      movej([-1.2302089344500047, -1.2969853503591224, -1.875639182904262, -1.539621866126728, 1.5731943360401213, -2.80099559440227], a=1.3962634015954636, v=1.0471975511965976)
    elif (32 == switch_1):
      $ 1983 "Case 32"
      $ 1985 "decap_Vial"
      $ 1986 "Set GRP_3F_Open=On"
      set_standard_digital_out(5, True)
      $ 1987 "MoveJ"
      $ 1988 "Waypoint_87" "breakAfter"
      movej(get_inverse_kin(Waypoint_87_p, qnear=Waypoint_87_q), a=0.5235987755982988, v=0.4363323129985824)
      $ 1989 "MoveL"
      $ 1990 "Vial_3FG_plac_1" "breakAfter"
      movel(Vial_3FG_plac_1_p, a=0.5, v=0.1)
      $ 1991 "Set GRP_3F_Open=Off"
      set_standard_digital_out(5, False)
      $ 1992 "Wait: 0.5"
      sleep(0.5)
      $ 1993 "MoveL"
      $ 1994 "Waypoint_88" "breakAfter"
      movel(Waypoint_88_p, a=0.5, v=0.1, r=0.05)
      $ 1995 "MoveJ"
      $ 1996 "cap_dump_1" "breakAfter"
      movej(get_inverse_kin(cap_dump_1_p, qnear=cap_dump_1_q), a=0.5235987755982988, v=0.4363323129985824)
      # begin: URCap Program Node
      #   Source: Robotiq_Grippers, 3.17.0.105337, Robotiq Inc.
      #   Type: Gripper
      $ 1997 "Gripper Open (1)"
      if not(gripper_connected[0]):
        popup("Gripper 1 must be connected to run this program.", "No connection", False, True, True)
      end
      if not(rq_is_gripper_activated("1")):
        popup("Gripper 1 is not activated. Go to Installation tab > Gripper to activate it and run the program again.", "Not activated", False, True, True)
      end
      rq_set_pos_spd_for(0, 255, 255, "1")
      rq_wait_pos_spe_for_request(0, 255, 255, "1")
      rq_go_to("1")
      rq_wait("1")
      # end: URCap Program Node
      $ 1998 "MoveJ"
      $ 1999 "Waypoint_89" "breakAfter"
      movej(get_inverse_kin(Waypoint_89_p, qnear=Waypoint_89_q), a=0.5235987755982988, v=0.4363323129985824, r=0.05)
      $ 2000 "MoveL"
      $ 2001 "Vial_3FG_plac_2" "breakAfter"
      movel(Vial_3FG_plac_2_p, a=0.5, v=0.1)
      # begin: URCap Program Node
      #   Source: Robotiq_Grippers, 3.17.0.105337, Robotiq Inc.
      #   Type: Gripper
      $ 2002 "Gripper Close (1)"
      if not(gripper_connected[0]):
        popup("Gripper 1 must be connected to run this program.", "No connection", False, True, True)
      end
      if not(rq_is_gripper_activated("1")):
        popup("Gripper 1 is not activated. Go to Installation tab > Gripper to activate it and run the program again.", "Not activated", False, True, True)
      end
      rq_set_pos_spd_for(255, 204, 255, "1")
      rq_wait_pos_spe_for_request(255, 204, 255, "1")
      rq_go_to("1")
      rq_wait("1")
      # end: URCap Program Node
      $ 2009 "Decap"
      $ 2010 "Action_Info≔'decapping'"
      global Action_Info="decapping"
      $ 2011 "Set GRP_3F_Enable=On"
      set_standard_digital_out(4, True)
      $ 2012 "Set GRP_3F_Decap=On"
      set_standard_digital_out(3, True)
      $ 2013 "Force"
      sleep(0.02)
      zero_ftsensor()
      force_mode(p[0.0,0.0,0.0,0.0,0.0,0.0], [0, 0, 1, 0, 0, 0], [0.0, 0.0, 1.0, 0.0, 0.0, 0.0], 2, [0.1, 0.1, 0.001, 0.3490658503988659, 0.3490658503988659, 0.3490658503988659])
      $ 2014 "check_decapping(offset=0.015, timeout=10, abort=CMD_Hold)" "noBreak"
      check_decapping(offset=0.015, timeout=10, abort=CMD_Hold)
      end_force_mode()
      stopl(5.0)
      $ 2015 "Set GRP_3F_Decap=Off"
      set_standard_digital_out(3, False)
      $ 2016 "Set GRP_3F_Enable=Off"
      set_standard_digital_out(4, False)
      $ 2017 "MoveL"
      $ 2018 "Waypoint_90" "breakAfter"
      movel(Waypoint_90_p, a=0.5, v=0.1, r=0.05)
      $ 2019 "MoveJ"
      $ 2020 "cap_dump_2" "breakAfter"
      movej(get_inverse_kin(cap_dump_2_p, qnear=cap_dump_2_q), a=0.5235987755982988, v=0.4363323129985824)
      # begin: URCap Program Node
      #   Source: Robotiq_Grippers, 3.17.0.105337, Robotiq Inc.
      #   Type: Gripper
      $ 2021 "Gripper Open (1)"
      if not(gripper_connected[0]):
        popup("Gripper 1 must be connected to run this program.", "No connection", False, True, True)
      end
      if not(rq_is_gripper_activated("1")):
        popup("Gripper 1 is not activated. Go to Installation tab > Gripper to activate it and run the program again.", "Not activated", False, True, True)
      end
      rq_set_pos_spd_for(0, 204, 255, "1")
      rq_wait_pos_spe_for_request(0, 204, 255, "1")
      rq_go_to("1")
      rq_wait("1")
      # end: URCap Program Node
      $ 2022 "MoveJ"
      $ 2023 "Waypoint_91" "breakAfter"
      movej(get_inverse_kin(Waypoint_91_p, qnear=Waypoint_91_q), a=0.5235987755982988, v=0.4363323129985824, r=0.036)
    elif (33 == switch_1):
      $ 2024 "Case 33"
      $ 2025 "Shake and liquid transfer"
      $ 2026 "MoveL"
      $ 2027 "Vial_liq_abov_1" "breakAfter"
      movel(Vial_liq_abov_1_p, a=0.5, v=0.1)
      $ 2028 "Vial_liq_pick_3" "breakAfter"
      movel(Vial_liq_pick_3_p, a=0.5, v=0.1)
      $ 2029 "Vial_liq_pick_4" "breakAfter"
      movel(Vial_liq_pick_4_p, a=0.5, v=0.1)
      # begin: URCap Program Node
      #   Source: Robotiq_Grippers, 3.17.0.105337, Robotiq Inc.
      #   Type: Gripper
      $ 2030 "Gripper Close (1)"
      if not(gripper_connected[0]):
        popup("Gripper 1 must be connected to run this program.", "No connection", False, True, True)
      end
      if not(rq_is_gripper_activated("1")):
        popup("Gripper 1 is not activated. Go to Installation tab > Gripper to activate it and run the program again.", "Not activated", False, True, True)
      end
      rq_set_pos_spd_for(255, 82, 71, "1")
      rq_wait_pos_spe_for_request(255, 82, 71, "1")
      rq_go_to("1")
      rq_wait("1")
      # end: URCap Program Node
      $ 2031 "Wait: 1.0"
      sleep(1.0)
      $ 2032 "Set GRP_3F_Open=On"
      set_standard_digital_out(5, True)
      $ 2033 "Wait: 0.5"
      sleep(0.5)
      $ 2034 "Vial_liq_abov_2" "breakAfter"
      movel(Vial_liq_abov_2_p, a=0.3, v=0.05, r=0.05)
      $ 2035 "MoveL"
      $ 2036 "Liquid_midway_1" "breakAfter"
      movel(Liquid_midway_1_p, a=0.5, v=0.1)
      $ 2037 "Loop 3 times"
      Loop_1 = 0
      while (Loop_1 < 3):
        $ 2038 "shake_3" "breakAfter"
        movel(shake_3_p, a=2.0, v=0.5)
        $ 2039 "shake_4" "breakAfter"
        movel(shake_4_p, a=2.0, v=0.5)
        Loop_1 = Loop_1 + 1
      end
      $ 2040 "drop_above_3" "breakAfter"
      movel(drop_above_3_p, a=0.5, v=0.1)
      $ 2041 "drop_above_4" "breakAfter"
      movel(drop_above_4_p, a=0.5, v=0.1)
      $ 2042 "liq_tran_3" "breakAfter"
      movel(liq_tran_3_p, a=0.5, v=0.05, r=0.008)
      $ 2043 "Wait: 1.0"
      sleep(1.0)
      $ 2044 "drop_above_5" "breakAfter"
      movel(drop_above_5_p, a=0.5, v=0.1)
      $ 2045 "Waypoint_92" "breakAfter"
      movel(Waypoint_92_p, a=0.5, v=0.1)
      $ 2046 "liq_tran_4" "breakAfter"
      movel(liq_tran_4_p, a=0.5, v=0.05)
      $ 2047 "Wait: 1.0"
      sleep(1.0)
      $ 2048 "drop_above_6" "breakAfter"
      movel(drop_above_6_p, a=0.5, v=0.1)
      $ 2049 "drop_above_7" "breakAfter"
      movel(drop_above_7_p, a=0.5, v=0.1)
      $ 2050 "Liquid_midway_2" "breakAfter"
      movel(Liquid_midway_2_p, a=0.5, v=0.1)
      $ 2051 "MoveL"
      $ 2052 "Vial_drop_abo_1" "breakAfter"
      movel(Vial_drop_abo_1_p, a=0.5, v=0.1)
      $ 2053 "Vial_liq_drop_1" "breakAfter"
      movel(Vial_liq_drop_1_p, a=0.5, v=0.1)
      # begin: URCap Program Node
      #   Source: Robotiq_Grippers, 3.17.0.105337, Robotiq Inc.
      #   Type: Gripper
      $ 2054 "Gripper Open (1)"
      if not(gripper_connected[0]):
        popup("Gripper 1 must be connected to run this program.", "No connection", False, True, True)
      end
      if not(rq_is_gripper_activated("1")):
        popup("Gripper 1 is not activated. Go to Installation tab > Gripper to activate it and run the program again.", "Not activated", False, True, True)
      end
      rq_set_pos_spd_for(0, 82, 71, "1")
      rq_wait_pos_spe_for_request(0, 82, 71, "1")
      rq_go_to("1")
      rq_wait("1")
      # end: URCap Program Node
      $ 2055 "Vial_drop_abo_2" "breakAfter"
      movel(Vial_drop_abo_2_p, a=0.5, v=0.1)
    elif (34 == switch_1):
      $ 2056 "Case 34"
      $ 2057 "Task≔'Dosing'"
      global Task="Dosing"
      $ 2058 "Powder dosing all"
      $ 2059 "send_target_info()"
      send_target_info()
      $ 2060 "zero_scale()"
      zero_scale()
      $ 2061 "prev_spat≔''"
      global prev_spat=""
      $ 2062 "spatula≔''"
      global spatula=""
      $ 2063 "send_powder_info()"
      send_powder_info()
      $ 2064 "Set AO[0]=0.0"
      set_standard_analog_out(0, 0.0)
      $ 2065 "Wait: 0.2"
      sleep(0.2)
      $ 2066 "reach pots decapping pose"
      # begin: URCap Program Node
      #   Source: SensoPart VISOR Robotic, 2.0.6, SensoPart Industriesensorik GmbH
      #   Type: VISOR Robotic App
      $ 2072 "VISOR Easy Pick"
      def visorFuncEasyPick_a93150():
        # begin: URCap Program Node
        #   Source: SensoPart VISOR Robotic, 2.0.6, SensoPart Industriesensorik GmbH
        #   Type: Easy Pick Setup
        $ 2073 "# 1 Setup" "noBreak"
        local easyPickVisorId = 1
        local easyPickArmMounted = True
        local easyPickSetJob = True
        local easyPickJobName = "Weight_scale"
        local easyPickAtImgAcq = False
        local easyPickImgAcqPose = Trigger
        # end: URCap Program Node
        # begin: URCap Program Node
        #   Source: SensoPart VISOR Robotic, 2.0.6, SensoPart Industriesensorik GmbH
        #   Type: Process
        $ 2074 "Process" "noBreak"
        local easyPickObjTaken = False
        local easyPickTrigger = False
        local easyPickPoseIdx = 0
        local easyPickPose = p[0,0,0,0,0,0]
        def easyPickFuncTrigger(visorId, setJob, jobName, arm):
        if (setJob):
          visor_changeJob(visorId, jobName, 6000)
        end
        if (arm):
          visor_trigger(visorId, 6000, "arm")
        else:
          visor_trigger(visorId, 6000)
        end
        global easyPickParts_4=visor_partsFound(visorId)
        visor_easyPickUpdate(visorId, "parts", visor_partsFound(visorId))
        return visor_getPose3d(visorId, 0)
      end
      while (not easyPickObjTaken):
        easyPickTrigger = (easyPickCount_4 >= visor_partsFound(easyPickVisorId)) or (easyPickCount_4 > 9) or (not visor_easyPickCheckIdent("3d2ec7", easyPickVisorId))
        if (easyPickTrigger):
          easyPickCount_4 = 0
        end
        easyPickPoseIdx = easyPickCount_4
        easyPickPose = visor_getPose3d(easyPickVisorId, easyPickPoseIdx)
        visor_easyPickUpdate(easyPickVisorId, "counter", easyPickPoseIdx)
        # begin: URCap Program Node
        #   Source: SensoPart VISOR Robotic, 2.0.6, SensoPart Industriesensorik GmbH
        #   Type: Image Acquisition Pose
        $ 2075 "Image Acquisition Pose" "noBreak"
        if (easyPickTrigger):
          if (not easyPickAtImgAcq):
            movej(pose_trans(easyPickImgAcqPose,p[0.0000,0.0000,-0.0000,0.0000,0.0000,0.0000]),a=1.3963,v=1.0472,t=0.000000,r=0.000000)
            easyPickAtImgAcq = True
          end
          easyPickPose = easyPickFuncTrigger(easyPickVisorId, easyPickSetJob, easyPickJobName, easyPickArmMounted)
        end
        # end: URCap Program Node
        # begin: URCap Program Node
        #   Source: SensoPart VISOR Robotic, 2.0.6, SensoPart Industriesensorik GmbH
        #   Type: Object Detected
        $ 2076 "Object Detected" "noBreak"
        if (visor_partsFound(easyPickVisorId) > 0):
          $ 2077 "Open Gripper" "noBreak"
          $ 2078 "weight_value≔get_weight()" "noBreak"
          global weight_value=get_weight()
          $ 2079 "Wait: 1.0" "noBreak"
          sleep(1.0)
          $ 2080 "diff≔target_weight-weight_value" "noBreak"
          global diff=target_weight-weight_value
          $ 2081 "compute_level_percent(W_now, weight_value)" "noBreak"
          compute_level_percent(W_now, weight_value)
          $ 2082 "send_level_info()" "noBreak"
          send_level_info()
          $ 2083 "spatula≔select_spatula(Flowability, level, diff, bulk_density, mouth_d)" "noBreak"
          global spatula=select_spatula(Flowability, level, diff, bulk_density, mouth_d)
          $ 2084 "Wait: 0.2" "noBreak"
          sleep(0.2)
          $ 2085 "send_spatula_info()" "noBreak"
          send_spatula_info()
          $ 2086 "If spatula ≟ 'spatula_L'" "noBreak"
          if (spatula  ==  "spatula_L"):
            $ 2087 "MoveJ" "noBreak"
            $ 2088 "Spatula_otw" "noBreak"
            movej(get_inverse_kin(Spatula_otw_p, qnear=Spatula_otw_q), a=1.3962634015954636, v=1.0471975511965976)
            $ 2089 "pick_spat_L_abv" "noBreak"
            movej(get_inverse_kin(pick_spat_L_abv_p, qnear=pick_spat_L_abv_q), a=1.3962634015954636, v=1.0471975511965976)
            $ 2090 "MoveL" "noBreak"
            $ 2091 "spat_L_pick" "noBreak"
            movel(spat_L_pick_p, a=1.2, v=0.25)
            # begin: URCap Program Node
            #   Source: Robotiq_Grippers, 3.17.0.105337, Robotiq Inc.
            #   Type: Gripper
            $ 2092 "Gripper Close (1)" "noBreak"
            if not(gripper_connected[0]):
              popup("Gripper 1 must be connected to run this program.", "No connection", False, True, True)
            end
            if not(rq_is_gripper_activated("1")):
              popup("Gripper 1 is not activated. Go to Installation tab > Gripper to activate it and run the program again.", "Not activated", False, True, True)
            end
            rq_set_pos_spd_for(255, 0, 77, "1")
            rq_wait_pos_spe_for_request(255, 0, 77, "1")
            rq_go_to("1")
            rq_wait("1")
            # end: URCap Program Node
            $ 2093 "spat_L_lift" "noBreak"
            movel(spat_L_lift_p, a=1.2, v=0.25, r=0.01)
            $ 2094 "spat_L_side" "noBreak"
            movel(spat_L_side_p, a=1.2, v=0.25, r=0.01)
            $ 2095 "spat_L_up" "noBreak"
            movel(spat_L_up_p, a=1.2, v=0.25, r=0.05)
            $ 2096 "MoveJ" "noBreak"
            $ 2097 "Spatula_otw" "noBreak"
            movej(get_inverse_kin(Spatula_otw_p, qnear=Spatula_otw_q), a=1.3962634015954636, v=1.0471975511965976)
          else:
            $ 2098 "ElseIf spatula ≟'spatula_M'" "noBreak"
            if (spatula  == "spatula_M"):
              $ 2099 "MoveJ" "noBreak"
              $ 2100 "Spatula_otw" "noBreak"
              movej(get_inverse_kin(Spatula_otw_p, qnear=Spatula_otw_q), a=1.3962634015954636, v=1.0471975511965976)
              $ 2101 "spat_M_up" "noBreak"
              movej(get_inverse_kin(spat_M_up_p, qnear=spat_M_up_q), a=1.3962634015954636, v=1.0471975511965976, r=0.05)
              $ 2102 "MoveL" "noBreak"
              $ 2103 "spat_M_pick" "noBreak"
              movel(spat_M_pick_p, a=1.2, v=0.25)
              # begin: URCap Program Node
              #   Source: Robotiq_Grippers, 3.17.0.105337, Robotiq Inc.
              #   Type: Gripper
              $ 2104 "Gripper Close (1)" "noBreak"
              if not(gripper_connected[0]):
                popup("Gripper 1 must be connected to run this program.", "No connection", False, True, True)
              end
              if not(rq_is_gripper_activated("1")):
                popup("Gripper 1 is not activated. Go to Installation tab > Gripper to activate it and run the program again.", "Not activated", False, True, True)
              end
              rq_set_pos_spd_for(255, 0, 77, "1")
              rq_wait_pos_spe_for_request(255, 0, 77, "1")
              rq_go_to("1")
              rq_wait("1")
              # end: URCap Program Node
              $ 2105 "spat_M_up" "noBreak"
              movel(spat_M_up_p, a=1.2, v=0.25, r=0.05)
              $ 2106 "Spatula_otw" "noBreak"
              movel(Spatula_otw_p, a=1.2, v=0.25)
              $ 2107 "switch_spat_M≔ False " "noBreak"
              global switch_spat_M=  False
            else:
              $ 2108 "ElseIf spatula≟'spatula_S'" "noBreak"
              if (spatula == "spatula_S"):
                $ 2109 "MoveJ" "noBreak"
                $ 2110 "Spatula_otw" "noBreak"
                movej(get_inverse_kin(Spatula_otw_p, qnear=Spatula_otw_q), a=1.3962634015954636, v=1.0471975511965976)
                $ 2111 "spat_S_Up_7" "noBreak"
                movej(get_inverse_kin(spat_S_Up_7_p, qnear=spat_S_Up_7_q), a=1.3962634015954636, v=1.0471975511965976, r=0.05)
                $ 2112 "MoveL" "noBreak"
                $ 2113 "spat_S_Pick_4" "noBreak"
                movel(spat_S_Pick_4_p, a=1.2, v=0.25)
                # begin: URCap Program Node
                #   Source: Robotiq_Grippers, 3.17.0.105337, Robotiq Inc.
                #   Type: Gripper
                $ 2114 "Gripper Close (1)" "noBreak"
                if not(gripper_connected[0]):
                  popup("Gripper 1 must be connected to run this program.", "No connection", False, True, True)
                end
                if not(rq_is_gripper_activated("1")):
                  popup("Gripper 1 is not activated. Go to Installation tab > Gripper to activate it and run the program again.", "Not activated", False, True, True)
                end
                rq_set_pos_spd_for(255, 0, 77, "1")
                rq_wait_pos_spe_for_request(255, 0, 77, "1")
                rq_go_to("1")
                rq_wait("1")
                # end: URCap Program Node
                $ 2115 "spat_S_Up_8" "noBreak"
                movel(spat_S_Up_8_p, a=1.2, v=0.25, r=0.05)
                $ 2116 "Spatula_otw" "noBreak"
                movel(Spatula_otw_p, a=1.2, v=0.25)
                $ 2117 "switch_spat_S≔ False " "noBreak"
                global switch_spat_S=  False
              else:
                $ 2118 "ElseIf spatula≟'spatula_flat_M'" "noBreak"
                if (spatula == "spatula_flat_M"):
                  $ 2119 "MoveJ" "noBreak"
                  $ 2120 "Spatula_otw" "noBreak"
                  movej(get_inverse_kin(Spatula_otw_p, qnear=Spatula_otw_q), a=1.3962634015954636, v=1.0471975511965976)
                  $ 2121 "spat_flatM_up" "noBreak"
                  movej(get_inverse_kin(spat_flatM_up_p, qnear=spat_flatM_up_q), a=1.3962634015954636, v=1.0471975511965976, r=0.05)
                  $ 2122 "MoveL" "noBreak"
                  $ 2123 "spat_flatM_pick" "noBreak"
                  movel(spat_flatM_pick_p, a=1.2, v=0.25)
                  # begin: URCap Program Node
                  #   Source: Robotiq_Grippers, 3.17.0.105337, Robotiq Inc.
                  #   Type: Gripper
                  $ 2124 "Gripper Close (1)" "noBreak"
                  if not(gripper_connected[0]):
                    popup("Gripper 1 must be connected to run this program.", "No connection", False, True, True)
                  end
                  if not(rq_is_gripper_activated("1")):
                    popup("Gripper 1 is not activated. Go to Installation tab > Gripper to activate it and run the program again.", "Not activated", False, True, True)
                  end
                  rq_set_pos_spd_for(255, 0, 77, "1")
                  rq_wait_pos_spe_for_request(255, 0, 77, "1")
                  rq_go_to("1")
                  rq_wait("1")
                  # end: URCap Program Node
                  $ 2125 "spat_flatM_up" "noBreak"
                  movel(spat_flatM_up_p, a=1.2, v=0.25, r=0.05)
                  $ 2126 "Spatula_otw" "noBreak"
                  movel(Spatula_otw_p, a=1.2, v=0.25)
                  $ 2127 "switch_spat_F_M≔ False " "noBreak"
                  global switch_spat_F_M=  False
                else:
                  $ 2128 "ElseIf spatula≟'spatula_flat_S'" "noBreak"
                  if (spatula == "spatula_flat_S"):
                    $ 2129 "MoveJ" "noBreak"
                    $ 2130 "Spatula_otw" "noBreak"
                    movej(get_inverse_kin(Spatula_otw_p, qnear=Spatula_otw_q), a=1.3962634015954636, v=1.0471975511965976)
                    $ 2131 "spat_flatS_up" "noBreak"
                    movej(get_inverse_kin(spat_flatS_up_p, qnear=spat_flatS_up_q), a=1.3962634015954636, v=1.0471975511965976, r=0.05)
                    $ 2132 "MoveL" "noBreak"
                    $ 2133 "spat_flatS_pick" "noBreak"
                    movel(spat_flatS_pick_p, a=1.2, v=0.25)
                    # begin: URCap Program Node
                    #   Source: Robotiq_Grippers, 3.17.0.105337, Robotiq Inc.
                    #   Type: Gripper
                    $ 2134 "Gripper Close (1)" "noBreak"
                    if not(gripper_connected[0]):
                      popup("Gripper 1 must be connected to run this program.", "No connection", False, True, True)
                    end
                    if not(rq_is_gripper_activated("1")):
                      popup("Gripper 1 is not activated. Go to Installation tab > Gripper to activate it and run the program again.", "Not activated", False, True, True)
                    end
                    rq_set_pos_spd_for(255, 0, 77, "1")
                    rq_wait_pos_spe_for_request(255, 0, 77, "1")
                    rq_go_to("1")
                    rq_wait("1")
                    # end: URCap Program Node
                    $ 2135 "spat_flatS_up" "noBreak"
                    movel(spat_flatS_up_p, a=1.2, v=0.25, r=0.05)
                    $ 2136 "Spatula_otw" "noBreak"
                    movel(Spatula_otw_p, a=1.2, v=0.25)
                    $ 2137 "switch_spat_F_S≔ False " "noBreak"
                    global switch_spat_F_S=  False
                  end
                end
              end
            end
          end
          $ 2138 "Action_Info≔'Scooping'" "noBreak"
          global Action_Info="Scooping"
          $ 2139 "auto_tilt_and_scoop(W_now, target_weight, weight_value)" "noBreak"
          auto_tilt_and_scoop(W_now, target_weight, weight_value)
          $ 2140 "Action_Info≔'Dosing'" "noBreak"
          global Action_Info="Dosing"
          # begin: URCap Program Node
          #   Source: SensoPart VISOR Robotic, 2.0.6, SensoPart Industriesensorik GmbH
          #   Type: Approach Pose
          $ 2141 "Approach Pose" "noBreak"
          movej(pose_trans(easyPickPose,p[0.0000,0.0000,-0.0000,0.0000,0.0000,0.0000]),a=0.2618,v=0.1745,t=0.000000,r=0.000000)
          # end: URCap Program Node
          # begin: URCap Program Node
          #   Source: SensoPart VISOR Robotic, 2.0.6, SensoPart Industriesensorik GmbH
          #   Type: Target Pose
          $ 2142 "Target Pose" "noBreak"
          movel(pose_trans(easyPickPose,p[0.0000,0.0000,-0.0000,0.0000,0.0000,0.0000]),a=0.0500,v=0.0200,t=0.000000,r=0.000000)
          # end: URCap Program Node
          $ 2143 "Close Gripper" "noBreak"
          $ 2144 "dispense_pos≔get_actual_tcp_pose()" "noBreak"
          global dispense_pos= get_actual_tcp_pose ()
          $ 2145 "Loop weight_value≤target_weight " "noBreak"
          thread Thread_while_2145():
            while (True):
              $ 2146 "MoveL" "noBreak"
              $ 2147 "dispense_pos" "noBreak"
              movel(dispense_pos, a=0.2, v=0.1)
              $ 2148 "log_weight()" "noBreak"
              log_weight()
              $ 2149 "If level≥85" "noBreak"
              if (level >= 85):
                $ 2150 "Rotate()" "noBreak"
                Rotate()
              end
              $ 2151 "If level≤85" "noBreak"
              if (level <= 85):
                $ 2152 "tilt_to_home()" "noBreak"
                tilt_to_home()
              end
              $ 2153 "Start_thread≔ True " "noBreak"
              global Start_thread=  True
              $ 2154 "vib_thread≔ True " "noBreak"
              global vib_thread=  True
              $ 2155 "Wait: 0.5" "noBreak"
              sleep(0.5)
              $ 2156 "If diff ≥(target_g*1.1)" "noBreak"
              if (diff  >= (target_g*1.1)):
                $ 2157 "tilt_pose≔pose_trans(get_actual_tcp_pose(), p[0, 0, 0, 0, 0, 2.0])" "noBreak"
                global tilt_pose=pose_trans(get_actual_tcp_pose(), p[0, 0, 0, 0, 0, 2.0])
                $ 2158 "movel(tilt_pose, a=0.5, v=0.5, r=0.00001)" "noBreak"
                movel(tilt_pose, a=0.5, v=0.5, r=0.00001)
              else:
                $ 2159 "Else" "noBreak"
                $ 2160 "Loop weight_value≤(target_weight-0.00) and tilt_angle≥(-1.999) and tilt_angle≤0.5" "noBreak"
                thread Thread_while_2160():
                  while (True):
                    $ 2161 "current_error≔target_weight-weight_value" "noBreak"
                    global current_error=target_weight-weight_value
                    $ 2162 "Integral_error≔Integral_error+current_error*dt" "noBreak"
                    global Integral_error=Integral_error+current_error*dt
                    $ 2163 "derivative≔(current_error-previous_error)/dt" "noBreak"
                    global derivative=(current_error-previous_error)/dt
                    $ 2164 "tilt_increment≔(kp*current_error)+(ki*Integral_error)+(kd*derivative)" "noBreak"
                    global tilt_increment=(kp*current_error)+(ki*Integral_error)+(kd*derivative)
                    $ 2165 "current_pose≔get_actual_tcp_pose()" "noBreak"
                    global current_pose= get_actual_tcp_pose ()
                    $ 2166 "tilt_angle≔current_pose[5]" "noBreak"
                    global tilt_angle=current_pose[5]
                    $ 2167 "tilt_pose≔pose_trans(current_pose, p[0, 0, 0, 0, 0, tilt_increment])" "noBreak"
                    global tilt_pose=pose_trans(current_pose, p[0, 0, 0, 0, 0, tilt_increment])
                    $ 2168 "movel(tilt_pose, a=0.3, v=0.3)" "noBreak"
                    movel(tilt_pose, a=0.3, v=0.3)
                    $ 2169 "previous_error≔current_error" "noBreak"
                    global previous_error=current_error
                  end
                end
                if (weight_value <= (target_weight-0.00)  and  tilt_angle >= (-1.999)  and  tilt_angle <= 0.5):
                  global thread_handler_2160=run Thread_while_2160()
                  while (weight_value <= (target_weight-0.00)  and  tilt_angle >= (-1.999)  and  tilt_angle <= 0.5):
                    sync()
                  end
                  kill thread_handler_2160
                end
              end
              $ 2170 "weight_value≔get_weight()" "noBreak"
              global weight_value=get_weight()
              $ 2172 "tilt_angle≔-1" "noBreak"
              global tilt_angle=-1
              $ 2173 "Wait: 0.5" "noBreak"
              sleep(0.5)
              $ 2174 "Start_thread≔ False " "noBreak"
              global Start_thread=  False
              $ 2175 "vib_thread≔ False " "noBreak"
              global vib_thread=  False
              $ 2177 "dispense_pos" "noBreak"
              movel(dispense_pos, a=1.2, v=0.25)
              $ 2178 "compute_level_percent(W_now, weight_value)" "noBreak"
              compute_level_percent(W_now, weight_value)
              $ 2179 "prev_spat≔spatula" "noBreak"
              global prev_spat=spatula
              $ 2180 "Wait: 0.2" "noBreak"
              sleep(0.2)
              $ 2181 "spatula≔select_spatula(Flowability, level, diff, bulk_density, mouth_d)" "noBreak"
              global spatula=select_spatula(Flowability, level, diff, bulk_density, mouth_d)
              $ 2182 "Wait: 1.0" "noBreak"
              sleep(1.0)
              $ 2183 "send_level_info()" "noBreak"
              send_level_info()
              $ 2184 "send_spatula_info()" "noBreak"
              send_spatula_info()
              $ 2185 "Integral_error≔0" "noBreak"
              global Integral_error=0
              $ 2186 "current_error≔0" "noBreak"
              global current_error=0
              $ 2187 "previous_error≔0" "noBreak"
              global previous_error=0
              $ 2188 "Set AO[0]=0.0" "noBreak"
              set_standard_analog_out(0, 0.0)
              $ 2189 "Wait: 0.5" "noBreak"
              sleep(0.5)
              $ 2190 "If spatula ≟ 'spatula_M' and switch_spat_M≟ True " "noBreak"
              if (spatula  ==  "spatula_M"  and  switch_spat_M ==   True  ):
                $ 2191 "MoveJ" "noBreak"
                $ 2192 "Spatula_otw" "noBreak"
                movej(get_inverse_kin(Spatula_otw_p, qnear=Spatula_otw_q), a=1.3962634015954636, v=1.0471975511965976)
                $ 2193 "spat_L_up" "noBreak"
                movej(get_inverse_kin(spat_L_up_p, qnear=spat_L_up_q), a=1.3962634015954636, v=1.0471975511965976)
                $ 2194 "MoveL" "noBreak"
                $ 2195 "spat_L_side" "noBreak"
                movel(spat_L_side_p, a=1.2, v=0.25)
                $ 2196 "spat_L_lift" "noBreak"
                movel(spat_L_lift_p, a=1.2, v=0.25)
                $ 2197 "spat_L_pick" "noBreak"
                movel(spat_L_pick_p, a=1.2, v=0.25)
                # begin: URCap Program Node
                #   Source: Robotiq_Grippers, 3.17.0.105337, Robotiq Inc.
                #   Type: Gripper
                $ 2198 "Gripper Open (1)" "noBreak"
                if not(gripper_connected[0]):
                  popup("Gripper 1 must be connected to run this program.", "No connection", False, True, True)
                end
                if not(rq_is_gripper_activated("1")):
                  popup("Gripper 1 is not activated. Go to Installation tab > Gripper to activate it and run the program again.", "Not activated", False, True, True)
                end
                rq_set_pos_spd_for(0, 255, 77, "1")
                rq_wait_pos_spe_for_request(0, 255, 77, "1")
                rq_go_to("1")
                rq_wait("1")
                # end: URCap Program Node
                $ 2199 "spat_M_pick" "noBreak"
                movel(spat_M_pick_p, a=1.2, v=0.25)
                # begin: URCap Program Node
                #   Source: Robotiq_Grippers, 3.17.0.105337, Robotiq Inc.
                #   Type: Gripper
                $ 2200 "Gripper Close (1)" "noBreak"
                if not(gripper_connected[0]):
                  popup("Gripper 1 must be connected to run this program.", "No connection", False, True, True)
                end
                if not(rq_is_gripper_activated("1")):
                  popup("Gripper 1 is not activated. Go to Installation tab > Gripper to activate it and run the program again.", "Not activated", False, True, True)
                end
                rq_set_pos_spd_for(255, 0, 77, "1")
                rq_wait_pos_spe_for_request(255, 0, 77, "1")
                rq_go_to("1")
                rq_wait("1")
                # end: URCap Program Node
                $ 2201 "spat_M_up" "noBreak"
                movel(spat_M_up_p, a=1.2, v=0.25)
                $ 2202 "Spatula_otw" "noBreak"
                movel(Spatula_otw_p, a=1.2, v=0.25)
                $ 2203 "switch_spat_M≔ False " "noBreak"
                global switch_spat_M=  False
              else:
                $ 2204 "ElseIf spatula ≟ 'spatula_S' and switch_spat_S ≟ True and prev_spat≟'spatula_M'" "noBreak"
                if (spatula  ==  "spatula_S" and switch_spat_S  ==   True  and prev_spat == "spatula_M"):
                  $ 2205 "MoveL" "noBreak"
                  $ 2206 "Spatula_otw" "noBreak"
                  movel(Spatula_otw_p, a=1.2, v=0.25)
                  $ 2207 "spat_M_up" "noBreak"
                  movel(spat_M_up_p, a=1.2, v=0.25)
                  $ 2208 "spat_M_pick" "noBreak"
                  movel(spat_M_pick_p, a=0.2, v=0.1)
                  # begin: URCap Program Node
                  #   Source: Robotiq_Grippers, 3.17.0.105337, Robotiq Inc.
                  #   Type: Gripper
                  $ 2209 "Gripper Open (1)" "noBreak"
                  if not(gripper_connected[0]):
                    popup("Gripper 1 must be connected to run this program.", "No connection", False, True, True)
                  end
                  if not(rq_is_gripper_activated("1")):
                    popup("Gripper 1 is not activated. Go to Installation tab > Gripper to activate it and run the program again.", "Not activated", False, True, True)
                  end
                  rq_set_pos_spd_for(0, 255, 77, "1")
                  rq_wait_pos_spe_for_request(0, 255, 77, "1")
                  rq_go_to("1")
                  rq_wait("1")
                  # end: URCap Program Node
                  $ 2210 "spat_S_pick" "noBreak"
                  movel(spat_S_pick_p, a=1.2, v=0.25)
                  # begin: URCap Program Node
                  #   Source: Robotiq_Grippers, 3.17.0.105337, Robotiq Inc.
                  #   Type: Gripper
                  $ 2211 "Gripper Close (1)" "noBreak"
                  if not(gripper_connected[0]):
                    popup("Gripper 1 must be connected to run this program.", "No connection", False, True, True)
                  end
                  if not(rq_is_gripper_activated("1")):
                    popup("Gripper 1 is not activated. Go to Installation tab > Gripper to activate it and run the program again.", "Not activated", False, True, True)
                  end
                  rq_set_pos_spd_for(255, 0, 77, "1")
                  rq_wait_pos_spe_for_request(255, 0, 77, "1")
                  rq_go_to("1")
                  rq_wait("1")
                  # end: URCap Program Node
                  $ 2212 "spat_S_up" "noBreak"
                  movel(spat_S_up_p, a=1.2, v=0.25)
                  $ 2213 "Spatula_otw" "noBreak"
                  movel(Spatula_otw_p, a=1.2, v=0.25)
                  $ 2214 "switch_spat_S≔ False " "noBreak"
                  global switch_spat_S=  False
                else:
                  $ 2215 "ElseIf spatula≟'spatula_S' and switch_spat_S≟ True  and prev_spat≟'spatula_L'" "noBreak"
                  if (spatula == "spatula_S" and switch_spat_S ==   True    and  prev_spat == "spatula_L"):
                    $ 2216 "MoveJ" "noBreak"
                    $ 2217 "Spatula_otw" "noBreak"
                    movej(get_inverse_kin(Spatula_otw_p, qnear=Spatula_otw_q), a=1.3962634015954636, v=1.0471975511965976)
                    $ 2218 "spat_L_up" "noBreak"
                    movej(get_inverse_kin(spat_L_up_p, qnear=spat_L_up_q), a=1.3962634015954636, v=1.0471975511965976)
                    $ 2219 "MoveL" "noBreak"
                    $ 2220 "spat_L_side" "noBreak"
                    movel(spat_L_side_p, a=1.2, v=0.25)
                    $ 2221 "spat_L_lift" "noBreak"
                    movel(spat_L_lift_p, a=1.2, v=0.25)
                    $ 2222 "spat_L_pick" "noBreak"
                    movel(spat_L_pick_p, a=0.25, v=0.15)
                    # begin: URCap Program Node
                    #   Source: Robotiq_Grippers, 3.17.0.105337, Robotiq Inc.
                    #   Type: Gripper
                    $ 2223 "Gripper Open (1)" "noBreak"
                    if not(gripper_connected[0]):
                      popup("Gripper 1 must be connected to run this program.", "No connection", False, True, True)
                    end
                    if not(rq_is_gripper_activated("1")):
                      popup("Gripper 1 is not activated. Go to Installation tab > Gripper to activate it and run the program again.", "Not activated", False, True, True)
                    end
                    rq_set_pos_spd_for(0, 255, 77, "1")
                    rq_wait_pos_spe_for_request(0, 255, 77, "1")
                    rq_go_to("1")
                    rq_wait("1")
                    # end: URCap Program Node
                    $ 2224 "spat_S_pick" "noBreak"
                    movel(spat_S_pick_p, a=1.2, v=0.25)
                    # begin: URCap Program Node
                    #   Source: Robotiq_Grippers, 3.17.0.105337, Robotiq Inc.
                    #   Type: Gripper
                    $ 2225 "Gripper Close (1)" "noBreak"
                    if not(gripper_connected[0]):
                      popup("Gripper 1 must be connected to run this program.", "No connection", False, True, True)
                    end
                    if not(rq_is_gripper_activated("1")):
                      popup("Gripper 1 is not activated. Go to Installation tab > Gripper to activate it and run the program again.", "Not activated", False, True, True)
                    end
                    rq_set_pos_spd_for(255, 0, 77, "1")
                    rq_wait_pos_spe_for_request(255, 0, 77, "1")
                    rq_go_to("1")
                    rq_wait("1")
                    # end: URCap Program Node
                    $ 2226 "spat_S_up" "noBreak"
                    movel(spat_S_up_p, a=1.2, v=0.25)
                    $ 2227 "Spatula_otw" "noBreak"
                    movel(Spatula_otw_p, a=1.2, v=0.25)
                    $ 2228 "switch_spat_S≔ False " "noBreak"
                    global switch_spat_S=  False
                  else:
                    $ 2229 "ElseIf spatula≟'spatula_flat_S'  and switch_spat_F_S ≟ True " "noBreak"
                    if (spatula == "spatula_flat_S"   and  switch_spat_F_S  ==   True  ):
                      $ 2230 "MoveL" "noBreak"
                      $ 2231 "Spatula_otw" "noBreak"
                      movel(Spatula_otw_p, a=1.2, v=0.25)
                      $ 2232 "spat_flatM_up" "noBreak"
                      movel(spat_flatM_up_p, a=1.2, v=0.25)
                      $ 2233 "spat_flatM_pick" "noBreak"
                      movel(spat_flatM_pick_p, a=1.2, v=0.25)
                      # begin: URCap Program Node
                      #   Source: Robotiq_Grippers, 3.17.0.105337, Robotiq Inc.
                      #   Type: Gripper
                      $ 2234 "Gripper Open (1)" "noBreak"
                      if not(gripper_connected[0]):
                        popup("Gripper 1 must be connected to run this program.", "No connection", False, True, True)
                      end
                      if not(rq_is_gripper_activated("1")):
                        popup("Gripper 1 is not activated. Go to Installation tab > Gripper to activate it and run the program again.", "Not activated", False, True, True)
                      end
                      rq_set_pos_spd_for(0, 0, 77, "1")
                      rq_wait_pos_spe_for_request(0, 0, 77, "1")
                      rq_go_to("1")
                      rq_wait("1")
                      # end: URCap Program Node
                      $ 2235 "spat_flatS_pick" "noBreak"
                      movel(spat_flatS_pick_p, a=1.2, v=0.25)
                      # begin: URCap Program Node
                      #   Source: Robotiq_Grippers, 3.17.0.105337, Robotiq Inc.
                      #   Type: Gripper
                      $ 2236 "Gripper Close (1)" "noBreak"
                      if not(gripper_connected[0]):
                        popup("Gripper 1 must be connected to run this program.", "No connection", False, True, True)
                      end
                      if not(rq_is_gripper_activated("1")):
                        popup("Gripper 1 is not activated. Go to Installation tab > Gripper to activate it and run the program again.", "Not activated", False, True, True)
                      end
                      rq_set_pos_spd_for(255, 0, 77, "1")
                      rq_wait_pos_spe_for_request(255, 0, 77, "1")
                      rq_go_to("1")
                      rq_wait("1")
                      # end: URCap Program Node
                      $ 2237 "spat_flatS_up" "noBreak"
                      movel(spat_flatS_up_p, a=1.2, v=0.25)
                      $ 2238 "Spatula_otw" "noBreak"
                      movel(Spatula_otw_p, a=1.2, v=0.25)
                      $ 2239 "switch_spat_F_S≔ False " "noBreak"
                      global switch_spat_F_S=  False
                    end
                  end
                end
              end
              $ 2240 "tilt(level)" "noBreak"
              tilt(level)
              $ 2241 "Action_Info≔'Scooping'" "noBreak"
              global Action_Info="Scooping"
              $ 2242 "auto_tilt_and_scoop(W_now, target_weight, weight_value)" "noBreak"
              auto_tilt_and_scoop(W_now, target_weight, weight_value)
              $ 2243 "Action_Info≔'Dosing'" "noBreak"
              global Action_Info="Dosing"
            end
          end
          if (weight_value <= target_weight ):
            global thread_handler_2145=run Thread_while_2145()
            while (weight_value <= target_weight ):
              sync()
            end
            kill thread_handler_2145
          end
          $ 2244 "Start_thread≔ False " "noBreak"
          global Start_thread=  False
          $ 2245 "vib_thread≔ False " "noBreak"
          global vib_thread=  False
          # begin: URCap Program Node
          #   Source: SensoPart VISOR Robotic, 2.0.6, SensoPart Industriesensorik GmbH
          #   Type: Exit Pose
          $ 2246 "Exit Pose" "noBreak"
          movel(pose_trans(easyPickPose,p[0.0000,0.0000,-0.0000,0.0000,0.0000,0.0000]),a=0.5000,v=0.2500,t=0.000000,r=0.000000)
          # end: URCap Program Node
          easyPickObjTaken = True
        end
        # end: URCap Program Node
        # begin: URCap Program Node
        #   Source: SensoPart VISOR Robotic, 2.0.6, SensoPart Industriesensorik GmbH
        #   Type: No Object Detected
        $ 2247 "No Object Detected" "noBreak"
        if (visor_partsFound(easyPickVisorId) < 1):
          $ 2248 "Popup: No weigh scale detected" "noBreak"
          popup("No weigh scale detected", "Message", False, False, blocking=True)
          else:
        end
        # end: URCap Program Node
      end
      easyPickCount_4 = easyPickCount_4 + 1
      visor_easyPickUpdate(easyPickVisorId, "counter", easyPickCount_4)
      visor_easyPickSetIdent("3d2ec7", easyPickVisorId)
      # end: URCap Program Node
    end
    visorFuncEasyPick_a93150()
    # end: URCap Program Node
    $ 2249 "MoveL"
    $ 2250 "dispense_pos" "breakAfter"
    movel(dispense_pos, a=0.2, v=0.1)
    $ 2251 "after_scoop()"
    after_scoop()
    $ 2252 "Place spatula back to the rack"
    $ 2253 "If spatula ≟ 'spatula_L'"
    if (spatula  ==  "spatula_L"):
      $ 2254 "MoveJ"
      $ 2255 "Spatula_otw" "breakAfter"
      movej(get_inverse_kin(Spatula_otw_p, qnear=Spatula_otw_q), a=1.3962634015954636, v=1.0471975511965976)
      $ 2256 "MoveL"
      $ 2257 "spat_L_up" "breakAfter"
      movel(spat_L_up_p, a=1.2, v=0.25, r=0.05)
      $ 2258 "spat_L_side" "breakAfter"
      movel(spat_L_side_p, a=1.2, v=0.25, r=0.01)
      $ 2259 "spat_L_lift" "breakAfter"
      movel(spat_L_lift_p, a=1.2, v=0.25, r=0.01)
      $ 2260 "spat_L_pick" "breakAfter"
      movel(spat_L_pick_p, a=0.25, v=0.15)
      # begin: URCap Program Node
      #   Source: Robotiq_Grippers, 3.17.0.105337, Robotiq Inc.
      #   Type: Gripper
      $ 2261 "Gripper Open (1)"
      if not(gripper_connected[0]):
        popup("Gripper 1 must be connected to run this program.", "No connection", False, True, True)
      end
      if not(rq_is_gripper_activated("1")):
        popup("Gripper 1 is not activated. Go to Installation tab > Gripper to activate it and run the program again.", "Not activated", False, True, True)
      end
      rq_set_pos_spd_for(0, 128, 128, "1")
      rq_wait_pos_spe_for_request(0, 128, 128, "1")
      rq_go_to("1")
      rq_wait("1")
      # end: URCap Program Node
      $ 2262 "MoveJ"
      $ 2263 "pick_spat_L_abv" "breakAfter"
      movej(get_inverse_kin(pick_spat_L_abv_p, qnear=pick_spat_L_abv_q), a=1.3962634015954636, v=1.0471975511965976)
      $ 2264 "Spatula_otw" "breakAfter"
      movej(get_inverse_kin(Spatula_otw_p, qnear=Spatula_otw_q), a=1.3962634015954636, v=1.0471975511965976)
    else:
      $ 2265 "ElseIf spatula ≟'spatula_M'"
      if (spatula  == "spatula_M"):
        $ 2266 "MoveJ"
        $ 2267 "Spatula_otw" "breakAfter"
        movej(get_inverse_kin(Spatula_otw_p, qnear=Spatula_otw_q), a=1.3962634015954636, v=1.0471975511965976)
        $ 2268 "spat_M_up" "breakAfter"
        movej(get_inverse_kin(spat_M_up_p, qnear=spat_M_up_q), a=1.3962634015954636, v=1.0471975511965976, r=0.05)
        $ 2269 "MoveL"
        $ 2270 "spat_M_pick" "breakAfter"
        movel(spat_M_pick_p, a=0.2, v=0.1)
        # begin: URCap Program Node
        #   Source: Robotiq_Grippers, 3.17.0.105337, Robotiq Inc.
        #   Type: Gripper
        $ 2271 "Gripper Open (1)"
        if not(gripper_connected[0]):
          popup("Gripper 1 must be connected to run this program.", "No connection", False, True, True)
        end
        if not(rq_is_gripper_activated("1")):
          popup("Gripper 1 is not activated. Go to Installation tab > Gripper to activate it and run the program again.", "Not activated", False, True, True)
        end
        rq_set_pos_spd_for(0, 128, 128, "1")
        rq_wait_pos_spe_for_request(0, 128, 128, "1")
        rq_go_to("1")
        rq_wait("1")
        # end: URCap Program Node
        $ 2272 "spat_M_up" "breakAfter"
        movel(spat_M_up_p, a=1.2, v=0.25, r=0.05)
        $ 2273 "Spatula_otw" "breakAfter"
        movel(Spatula_otw_p, a=1.2, v=0.25)
        $ 2274 "switch_spat_M≔ False "
        global switch_spat_M=  False
      else:
        $ 2275 "ElseIf spatula≟'spatula_S'"
        if (spatula == "spatula_S"):
          $ 2276 "MoveJ"
          $ 2277 "Spatula_otw" "breakAfter"
          movej(get_inverse_kin(Spatula_otw_p, qnear=Spatula_otw_q), a=1.3962634015954636, v=1.0471975511965976)
          $ 2278 "spat_S_Up_7" "breakAfter"
          movej(get_inverse_kin(spat_S_Up_7_p, qnear=spat_S_Up_7_q), a=1.3962634015954636, v=1.0471975511965976, r=0.05)
          $ 2279 "MoveL"
          $ 2280 "spat_S_Pick_4" "breakAfter"
          movel(spat_S_Pick_4_p, a=0.2, v=0.1)
          # begin: URCap Program Node
          #   Source: Robotiq_Grippers, 3.17.0.105337, Robotiq Inc.
          #   Type: Gripper
          $ 2281 "Gripper Open (1)"
          if not(gripper_connected[0]):
            popup("Gripper 1 must be connected to run this program.", "No connection", False, True, True)
          end
          if not(rq_is_gripper_activated("1")):
            popup("Gripper 1 is not activated. Go to Installation tab > Gripper to activate it and run the program again.", "Not activated", False, True, True)
          end
          rq_set_pos_spd_for(0, 255, 51, "1")
          rq_wait_pos_spe_for_request(0, 255, 51, "1")
          rq_go_to("1")
          rq_wait("1")
          # end: URCap Program Node
          $ 2282 "spat_S_Up_8" "breakAfter"
          movel(spat_S_Up_8_p, a=1.2, v=0.25, r=0.05)
          $ 2283 "Spatula_otw" "breakAfter"
          movel(Spatula_otw_p, a=1.2, v=0.25)
          $ 2284 "switch_spat_S≔ False "
          global switch_spat_S=  False
        else:
          $ 2285 "ElseIf spatula≟'spatula_flat_M'"
          if (spatula == "spatula_flat_M"):
            $ 2286 "MoveJ"
            $ 2287 "Spatula_otw" "breakAfter"
            movej(get_inverse_kin(Spatula_otw_p, qnear=Spatula_otw_q), a=1.3962634015954636, v=1.0471975511965976)
            $ 2288 "spat_flatM_up" "breakAfter"
            movej(get_inverse_kin(spat_flatM_up_p, qnear=spat_flatM_up_q), a=1.3962634015954636, v=1.0471975511965976, r=0.05)
            $ 2289 "MoveL"
            $ 2290 "spat_flatM_pick" "breakAfter"
            movel(spat_flatM_pick_p, a=1.2, v=0.25)
            # begin: URCap Program Node
            #   Source: Robotiq_Grippers, 3.17.0.105337, Robotiq Inc.
            #   Type: Gripper
            $ 2291 "Gripper Open (1)"
            if not(gripper_connected[0]):
              popup("Gripper 1 must be connected to run this program.", "No connection", False, True, True)
            end
            if not(rq_is_gripper_activated("1")):
              popup("Gripper 1 is not activated. Go to Installation tab > Gripper to activate it and run the program again.", "Not activated", False, True, True)
            end
            rq_set_pos_spd_for(0, 128, 128, "1")
            rq_wait_pos_spe_for_request(0, 128, 128, "1")
            rq_go_to("1")
            rq_wait("1")
            # end: URCap Program Node
            $ 2292 "spat_flatM_up" "breakAfter"
            movel(spat_flatM_up_p, a=1.2, v=0.25, r=0.05)
            $ 2293 "Spatula_otw" "breakAfter"
            movel(Spatula_otw_p, a=1.2, v=0.25)
            $ 2294 "switch_spat_F_M≔ False "
            global switch_spat_F_M=  False
          else:
            $ 2295 "ElseIf spatula≟'spatula_flat_S'"
            if (spatula == "spatula_flat_S"):
              $ 2296 "MoveJ"
              $ 2297 "Spatula_otw" "breakAfter"
              movej(get_inverse_kin(Spatula_otw_p, qnear=Spatula_otw_q), a=1.3962634015954636, v=1.0471975511965976)
              $ 2298 "spat_flatS_up" "breakAfter"
              movej(get_inverse_kin(spat_flatS_up_p, qnear=spat_flatS_up_q), a=1.3962634015954636, v=1.0471975511965976, r=0.05)
              $ 2299 "MoveL"
              $ 2300 "spat_flatS_pick" "breakAfter"
              movel(spat_flatS_pick_p, a=1.2, v=0.25)
              # begin: URCap Program Node
              #   Source: Robotiq_Grippers, 3.17.0.105337, Robotiq Inc.
              #   Type: Gripper
              $ 2301 "Gripper Open (1)"
              if not(gripper_connected[0]):
                popup("Gripper 1 must be connected to run this program.", "No connection", False, True, True)
              end
              if not(rq_is_gripper_activated("1")):
                popup("Gripper 1 is not activated. Go to Installation tab > Gripper to activate it and run the program again.", "Not activated", False, True, True)
              end
              rq_set_pos_spd_for(0, 128, 128, "1")
              rq_wait_pos_spe_for_request(0, 128, 128, "1")
              rq_go_to("1")
              rq_wait("1")
              # end: URCap Program Node
              $ 2302 "spat_flatS_up" "breakAfter"
              movel(spat_flatS_up_p, a=1.2, v=0.25, r=0.05)
              $ 2303 "Spatula_otw" "breakAfter"
              movel(Spatula_otw_p, a=1.2, v=0.25)
              $ 2304 "switch_spat_F_S≔ False "
              global switch_spat_F_S=  False
            end
          end
        end
      end
    end
    $ 2305 "switch_spat_M≔ True "
    global switch_spat_M=  True
    $ 2306 "switch_spat_S≔ True "
    global switch_spat_S=  True
    $ 2307 "switch_spat_F_M≔ True "
    global switch_spat_F_M=  True
    $ 2308 "switch_spat_F_S≔ True "
    global switch_spat_F_S=  True
    $ 2309 "Pick container from PoTS"
    $ 2310 "cont_place_offs≔pose_add(container_place, p[0.05,0,0,0,0,0])"
    global cont_place_offs=pose_add(container_place, p[0.05,0,0,0,0,0])
    $ 2311 "MoveJ"
    $ 2312 "cont_place_offs" "breakAfter"
    movej(cont_place_offs, a=1.3962634015954636, v=1.0471975511965976)
    $ 2313 "container_place" "breakAfter"
    movej(container_place, a=1.3962634015954636, v=1.0471975511965976)
    $ 2314 "MoveL"
    $ 2315 "target_pose" "breakAfter"
    movel(target_pose, a=1.2, v=0.25)
    # begin: URCap Program Node
    #   Source: Robotiq_Grippers, 3.17.0.105337, Robotiq Inc.
    #   Type: Gripper
    $ 2316 "Gripper Close (1)"
    if not(gripper_connected[0]):
      popup("Gripper 1 must be connected to run this program.", "No connection", False, True, True)
    end
    if not(rq_is_gripper_activated("1")):
      popup("Gripper 1 is not activated. Go to Installation tab > Gripper to activate it and run the program again.", "Not activated", False, True, True)
    end
    rq_set_pos_spd_for(255, 77, 77, "1")
    rq_wait_pos_spe_for_request(255, 77, 77, "1")
    rq_go_to("1")
    rq_wait("1")
    # end: URCap Program Node
    $ 2317 "container_place" "breakAfter"
    movel(container_place, a=0.6, v=0.1)
  elif (38 == switch_1):
    $ 2629 "Case 38"
    $ 2630 "Decap Powder container"
    $ 2631 "MoveJ"
    $ 2633 "Waypoint_7" "breakAfter"
    movej(get_inverse_kin(Waypoint_7_p, qnear=Waypoint_7_q), a=1.3962634015954636, v=1.0471975511965976, r=0.05)
    $ 2634 "MoveL"
    $ 2636 "Waypoint_8" "breakAfter"
    movel(Waypoint_8_p, a=1.2, v=0.25)
    $ 2637 "MoveL"
    $ 2638 "Decapp_above_3" "breakAfter"
    movel(Decapp_above_3_p, a=1.2, v=0.25)
    $ 2639 "Set GRP_3F_Open=On"
    set_standard_digital_out(5, True)
    $ 2640 "Wait: 0.5"
    sleep(0.5)
    $ 2641 "Decapp_place_3" "breakAfter"
    movel(Decapp_place_3_p, a=0.3, v=0.05)
    $ 2642 "Set GRP_3F_Open=Off"
    set_standard_digital_out(5, False)
    $ 2643 "Wait: 0.5"
    sleep(0.5)
    # begin: URCap Program Node
    #   Source: Robotiq_Grippers, 3.17.0.105337, Robotiq Inc.
    #   Type: Gripper
    $ 2644 "Gripper Open (1)"
    if not(gripper_connected[0]):
      popup("Gripper 1 must be connected to run this program.", "No connection", False, True, True)
    end
    if not(rq_is_gripper_activated("1")):
      popup("Gripper 1 is not activated. Go to Installation tab > Gripper to activate it and run the program again.", "Not activated", False, True, True)
    end
    rq_set_pos_spd_for(0, 77, 77, "1")
    rq_wait_pos_spe_for_request(0, 77, 77, "1")
    rq_go_to("1")
    rq_wait("1")
    # end: URCap Program Node
    $ 2645 "MoveL"
    $ 2646 "Decapp_above_4" "breakAfter"
    movel(Decapp_above_4_p, a=1.2, v=0.25)
    $ 2647 "Waypoint_78" "breakAfter"
    movel(Waypoint_78_p, a=1.2, v=0.25, r=0.05)
    $ 2648 "Home (Safe)"
    movej([-1.2302089344500047, -1.2969853503591224, -1.875639182904262, -1.539621866126728, 1.5731943360401213, -2.80099559440227], a=1.3962634015954636, v=1.0471975511965976)
  elif (39 == switch_1):
    $ 2649 "Case 39"
    $ 2650 "Powder container Pick"
    $ 2651 "Direct Pick"
    $ 2652 "Set"
    set_tcp(p[0.0,0.0,0.15052000000000001,3.1415,0.0,0.0])
    $ 2653 "read_db_data()"
    read_db_data()
    # begin: URCap Program Node
    #   Source: SensoPart VISOR Robotic, 2.0.6, SensoPart Industriesensorik GmbH
    #   Type: VISOR ChangeJob
    $ 2654 "# 1 VISOR ChangeJob"
    visor_changeJob(1, "Aztec_no_dot_pick", 6000)
    # end: URCap Program Node
    # begin: URCap Program Node
    #   Source: SensoPart VISOR Robotic, 2.0.6, SensoPart Industriesensorik GmbH
    #   Type: VISOR Terminal
    $ 2655 "# 1 VISOR Terminal"
    visor_terminal(1, "TRX00", 3000)
    # end: URCap Program Node
    $ 2656 "table_pick_TCP≔visor_getPose3d(1, 0)"
    global table_pick_TCP= visor_getPose3d (1, 0)
    # begin: URCap Program Node
    #   Source: Robotiq_Grippers, 3.17.0.105337, Robotiq Inc.
    #   Type: Gripper
    $ 2657 "Gripper Open (1)"
    if not(gripper_connected[0]):
      popup("Gripper 1 must be connected to run this program.", "No connection", False, True, True)
    end
    if not(rq_is_gripper_activated("1")):
      popup("Gripper 1 is not activated. Go to Installation tab > Gripper to activate it and run the program again.", "Not activated", False, True, True)
    end
    rq_set_pos_spd_for(0, 77, 77, "1")
    rq_wait_pos_spe_for_request(0, 77, 77, "1")
    rq_go_to("1")
    rq_wait("1")
    # end: URCap Program Node
    $ 2658 "MoveJ"
    $ 2660 "Waypoint_10" "breakAfter"
    movej(get_inverse_kin(Waypoint_10_p, qnear=Waypoint_10_q), a=1.3962634015954636, v=1.0471975511965976, r=0.05)
    $ 2661 "Waypoint_9" "breakAfter"
    movej(get_inverse_kin(Waypoint_9_p, qnear=Waypoint_9_q), a=1.3962634015954636, v=1.0471975511965976, r=0.05)
    $ 2662 "MoveJ"
    $ 2663 "table_pick_TCP" "breakAfter"
    movej(table_pick_TCP, a=0.8726646259971648, v=0.6981317007977318)
    $ 2664 "table_prepick≔pose_trans(table_pick_TCP,p[0,0,cent_edge/2,0,0,0])"
    global table_prepick=pose_trans(table_pick_TCP,p[0,0,cent_edge/2,0,0,0])
    $ 2665 "table_prepick" "breakAfter"
    movej(table_prepick, a=0.8726646259971648, v=0.6981317007977318)
    $ 2666 "table_safe_pick≔pose_trans(table_prepick, p[0,pick_2_base-H_c,cent_edge/2,0,0,0])"
    global table_safe_pick= pose_trans (table_prepick, p[0,pick_2_base-H_c,cent_edge/2,0,0,0])
    $ 2667 "table_safe_pick" "breakAfter"
    movej(table_safe_pick, a=0.8726646259971648, v=0.6981317007977318, r=0.05)
    $ 2668 "table_pick≔pose_trans(table_prepick, p[0,pick_2_base - d_cc,0,0,0,0])"
    global table_pick= pose_trans (table_prepick, p[0,pick_2_base - d_cc,0,0,0,0])
    $ 2669 "table_pick" "breakAfter"
    movej(table_pick, a=0.8726646259971648, v=0.6981317007977318)
    # begin: URCap Program Node
    #   Source: Robotiq_Grippers, 3.17.0.105337, Robotiq Inc.
    #   Type: Gripper
    $ 2670 "Gripper Close (1)"
    if not(gripper_connected[0]):
      popup("Gripper 1 must be connected to run this program.", "No connection", False, True, True)
    end
    if not(rq_is_gripper_activated("1")):
      popup("Gripper 1 is not activated. Go to Installation tab > Gripper to activate it and run the program again.", "Not activated", False, True, True)
    end
    rq_set_pos_spd_for(255, 77, 51, "1")
    rq_wait_pos_spe_for_request(255, 77, 51, "1")
    rq_go_to("1")
    rq_wait("1")
    # end: URCap Program Node
    $ 2671 "table_prepick" "breakAfter"
    movej(table_prepick, a=0.8726646259971648, v=0.6981317007977318)
    $ 2701 "powder_position≔'Position2'"
    global powder_position="Position2"
    $ 2702 "MoveJ"
    $ 2703 "Powder_wayp1" "breakAfter"
    movej(get_inverse_kin(Powder_wayp1_p, qnear=Powder_wayp1_q), a=1.3962634015954636, v=1.0471975511965976, r=0.05)
    $ 2704 "MoveL"
    $ 2705 "Waypoint_2" "breakAfter"
    movel(Waypoint_2_p, a=1.2, v=0.25)
    $ 2706 "Set"
    set_tcp(p[0.0,0.0,0.161,3.1415,0.0,0.0])
    $ 2707 "If powder_position ≟ 'Position1'"
    if (powder_position  ==  "Position1"):
      $ 2708 "MoveJ"
      $ 2709 "Postions_otw" "breakAfter"
      movej(get_inverse_kin(Postions_otw_p, qnear=Postions_otw_q), a=1.3962634015954636, v=1.0471975511965976, r=0.01)
      $ 2710 "MoveL"
      $ 2711 "Cont_A_TCP" "breakAfter"
      movel(Cont_A_TCP, a=0.5, v=0.2)
      $ 2712 "cont_A_prepick≔pose_trans(Cont_A_TCP, p[0,0,cent_edge/2,0,0,0])"
      global cont_A_prepick= pose_trans (Cont_A_TCP, p[0,0,cent_edge/2,0,0,0])
      $ 2713 "cont_A_prepick" "breakAfter"
      movel(cont_A_prepick, a=0.3, v=0.05)
      $ 2714 "cont_A_pick≔pose_trans(cont_A_prepick, p[0,pick_2_base-d_cc,0,0,0,0])"
      global cont_A_pick= pose_trans (cont_A_prepick, p[0,pick_2_base-d_cc,0,0,0,0])
      $ 2715 "cont_A_pick" "breakAfter"
      movel(cont_A_pick, a=0.2, v=0.1)
      # begin: URCap Program Node
      #   Source: Robotiq_Grippers, 3.17.0.105337, Robotiq Inc.
      #   Type: Gripper
      $ 2716 "Gripper Open (1)"
      if not(gripper_connected[0]):
        popup("Gripper 1 must be connected to run this program.", "No connection", False, True, True)
      end
      if not(rq_is_gripper_activated("1")):
        popup("Gripper 1 is not activated. Go to Installation tab > Gripper to activate it and run the program again.", "Not activated", False, True, True)
      end
      rq_set_pos_spd_for(0, 77, 26, "1")
      rq_wait_pos_spe_for_request(0, 77, 26, "1")
      rq_go_to("1")
      rq_wait("1")
      # end: URCap Program Node
      $ 2717 "cont_A_otw" "breakAfter"
      movel(cont_A_otw_p, a=0.5, v=0.2)
      $ 2718 "cont_A_prepick" "breakAfter"
      movel(cont_A_prepick, a=0.5, v=0.2)
      $ 2719 "Postions_otw" "breakAfter"
      movel(Postions_otw_p, a=0.5, v=0.2, r=0.01)
      $ 2721 "Home (Safe)"
      movej([-1.2302089344500047, -1.2969853503591224, -1.875639182904262, -1.539621866126728, 1.5731943360401213, -2.80099559440227], a=1.3962634015954636, v=1.0471975511965976)
    else:
      $ 2723 "ElseIf powder_position≟'Position2'"
      if (powder_position == "Position2"):
        $ 2724 "MoveJ"
        $ 2725 "Postions_otw" "breakAfter"
        movej(get_inverse_kin(Postions_otw_p, qnear=Postions_otw_q), a=1.3962634015954636, v=1.0471975511965976, r=0.01)
        $ 2726 "MoveL"
        $ 2729 "cont_B_prepick≔pose_trans(Cont_B_TCP, p[0,0,cent_edge/2,0,0,0])"
        global cont_B_prepick= pose_trans (Cont_B_TCP, p[0,0,cent_edge/2,0,0,0])
        $ 2730 "cont_B_prepick" "breakAfter"
        movel(cont_B_prepick, a=0.3, v=0.05)
        $ 2731 "cont_B_pick≔pose_trans(cont_B_prepick, p[0,pick_2_base-d_cc,0,0,0,0])"
        global cont_B_pick= pose_trans (cont_B_prepick, p[0,pick_2_base-d_cc,0,0,0,0])
        $ 2732 "cont_B_pick" "breakAfter"
        global move_thread_flag_2732=0
        thread move_thread_2732():
          enter_critical
          move_thread_flag_2732 = 1
          movel(cont_B_pick, a=0.2, v=0.1)
          move_thread_flag_2732 = 2
          exit_critical
        end
        move_thread_flag_2732 = 0
        move_thread_han_2732 = run move_thread_2732()
        while (True):
          local targetTcpDirection=get_target_tcp_speed()
          local stepsToRetract=tool_contact(direction=targetTcpDirection, force_threshold=8.000000)
          if (stepsToRetract > 0):
            kill move_thread_han_2732
            stopl(3.0)
            local backTrackMovement=get_actual_joint_positions_history(stepsToRetract)
            local contactPose=get_forward_kin(backTrackMovement)
            local posDir=[targetTcpDirection[0],targetTcpDirection[1],targetTcpDirection[2]]
            local retractTo=contactPose
            if (norm(posDir) > 1e-6):
              local normalizedPosDir=normalize(posDir)
              local additionalRetraction=p[normalizedPosDir[0] * 0.0, normalizedPosDir[1] * 0.0, normalizedPosDir[2] * 0.0, 0, 0, 0]
              retractTo = pose_sub(contactPose, additionalRetraction)
            end
            movel(retractTo, a=3.0, v=0.1)
            $ 2733 "Until (tool_contact_detection)"
            $ 2734 "saved_place_pos≔get_actual_tcp_pose()"
            global saved_place_pos= get_actual_tcp_pose ()
            break
          end
          sleep(1.0E-10)
          if (move_thread_flag_2732 > 1):
            join move_thread_han_2732
            break
          end
          sync()
        end
        # begin: URCap Program Node
        #   Source: Robotiq_Grippers, 3.17.0.105337, Robotiq Inc.
        #   Type: Gripper
        $ 2735 "Gripper Open (1)"
        if not(gripper_connected[0]):
          popup("Gripper 1 must be connected to run this program.", "No connection", False, True, True)
        end
        if not(rq_is_gripper_activated("1")):
          popup("Gripper 1 is not activated. Go to Installation tab > Gripper to activate it and run the program again.", "Not activated", False, True, True)
        end
        rq_set_pos_spd_for(0, 77, 26, "1")
        rq_wait_pos_spe_for_request(0, 77, 26, "1")
        rq_go_to("1")
        rq_wait("1")
        # end: URCap Program Node
        $ 2736 "cont_B_otw" "breakAfter"
        movel(cont_B_otw_p, a=1.2, v=0.25)
        $ 2738 "cont_B_safe" "breakAfter"
        movel(cont_B_safe_p, a=1.2, v=0.25)
        $ 2739 "Postions_otw" "breakAfter"
        movel(Postions_otw_p, a=1.2, v=0.25)
        $ 2741 "Home (Safe)"
        movej([-1.2302089344500047, -1.2969853503591224, -1.875639182904262, -1.539621866126728, 1.5731943360401213, -2.80099559440227], a=1.3962634015954636, v=1.0471975511965976)
      else:
        $ 2743 "ElseIf powder_position≟'Position3'"
        if (powder_position == "Position3"):
          $ 2744 "MoveJ"
          $ 2745 "Postions_otw" "breakAfter"
          movej(get_inverse_kin(Postions_otw_p, qnear=Postions_otw_q), a=1.3962634015954636, v=1.0471975511965976, r=0.01)
          $ 2752 "MoveL"
          $ 2753 "Cont_C_TCP" "breakAfter"
          movel(Cont_C_TCP, a=1.2, v=0.25, r=0.01)
          $ 2754 "cont_C_prepick≔pose_trans(Cont_C_TCP, p[0,0,cent_edge/2,0,0,0])"
          global cont_C_prepick= pose_trans (Cont_C_TCP, p[0,0,cent_edge/2,0,0,0])
          $ 2755 "cont_C_prepick" "breakAfter"
          movel(cont_C_prepick, a=0.3, v=0.05)
          $ 2756 "cont_C_pick≔pose_trans(cont_C_prepick, p[0,pick_2_base-d_cc,0,0,0,0])"
          global cont_C_pick= pose_trans (cont_C_prepick, p[0,pick_2_base-d_cc,0,0,0,0])
          $ 2757 "cont_C_pick" "breakAfter"
          movel(cont_C_pick, a=0.2, v=0.1)
          # begin: URCap Program Node
          #   Source: Robotiq_Grippers, 3.17.0.105337, Robotiq Inc.
          #   Type: Gripper
          $ 2758 "Gripper Open (1)"
          if not(gripper_connected[0]):
            popup("Gripper 1 must be connected to run this program.", "No connection", False, True, True)
          end
          if not(rq_is_gripper_activated("1")):
            popup("Gripper 1 is not activated. Go to Installation tab > Gripper to activate it and run the program again.", "Not activated", False, True, True)
          end
          rq_set_pos_spd_for(0, 77, 26, "1")
          rq_wait_pos_spe_for_request(0, 77, 26, "1")
          rq_go_to("1")
          rq_wait("1")
          # end: URCap Program Node
          $ 2759 "cont_C_otw" "breakAfter"
          movel(cont_C_otw_p, a=1.2, v=0.25)
          $ 2760 "cont_C_prepick" "breakAfter"
          movel(cont_C_prepick, a=1.2, v=0.25, r=0.01)
          $ 2761 "Postions_otw" "breakAfter"
          movel(Postions_otw_p, a=1.2, v=0.25)
          $ 2762 "Home (Safe)"
          movej([-1.2302089344500047, -1.2969853503591224, -1.875639182904262, -1.539621866126728, 1.5731943360401213, -2.80099559440227], a=1.3962634015954636, v=1.0471975511965976)
        end
      end
    end
    $ 2775 "Home (Safe)"
    movej([-1.2302089344500047, -1.2969853503591224, -1.875639182904262, -1.539621866126728, 1.5731943360401213, -2.80099559440227], a=1.3962634015954636, v=1.0471975511965976)
  elif (41 == switch_1):
    $ 2884 "Case 41"
    $ 2885 "Task≔'Decapping'"
    global Task="Decapping"
    $ 2886 "Weigh, Place & decap container"
    $ 2887 "Set"
    set_tcp(p[0.0,0.0,0.15052000000000001,3.1415,0.0,0.0])
    # begin: URCap Program Node
    #   Source: SensoPart VISOR Robotic, 2.0.6, SensoPart Industriesensorik GmbH
    #   Type: VISOR Robotic App
    $ 2888 "VISOR Easy Pick"
    def visorFuncEasyPick_316065():
      # begin: URCap Program Node
      #   Source: SensoPart VISOR Robotic, 2.0.6, SensoPart Industriesensorik GmbH
      #   Type: Easy Pick Setup
      $ 2889 "# 1 Setup" "noBreak"
      local easyPickVisorId = 1
      local easyPickArmMounted = True
      local easyPickSetJob = True
      local easyPickJobName = "PoTS"
      local easyPickAtImgAcq = False
      local easyPickImgAcqPose = FRM_PoTS
      # end: URCap Program Node
      # begin: URCap Program Node
      #   Source: SensoPart VISOR Robotic, 2.0.6, SensoPart Industriesensorik GmbH
      #   Type: Process
      $ 2890 "Process" "noBreak"
      local easyPickObjTaken = False
      local easyPickTrigger = False
      local easyPickPoseIdx = 0
      local easyPickPose = p[0,0,0,0,0,0]
      def easyPickFuncTrigger(visorId, setJob, jobName, arm):
      if (setJob):
        visor_changeJob(visorId, jobName, 6000)
      end
      if (arm):
        visor_trigger(visorId, 6000, "arm")
      else:
        visor_trigger(visorId, 6000)
      end
      global easyPickParts_7=visor_partsFound(visorId)
      visor_easyPickUpdate(visorId, "parts", visor_partsFound(visorId))
      return visor_getPose3d(visorId, 0)
    end
    while (not easyPickObjTaken):
      easyPickTrigger = (easyPickCount_7 >= visor_partsFound(easyPickVisorId)) or (easyPickCount_7 > 9) or (not visor_easyPickCheckIdent("133617", easyPickVisorId))
      if (easyPickTrigger):
        easyPickCount_7 = 0
      end
      easyPickPoseIdx = easyPickCount_7
      easyPickPose = visor_getPose3d(easyPickVisorId, easyPickPoseIdx)
      visor_easyPickUpdate(easyPickVisorId, "counter", easyPickPoseIdx)
      # begin: URCap Program Node
      #   Source: SensoPart VISOR Robotic, 2.0.6, SensoPart Industriesensorik GmbH
      #   Type: Image Acquisition Pose
      $ 2891 "Image Acquisition Pose" "noBreak"
      if (easyPickTrigger):
        if (not easyPickAtImgAcq):
          movej(pose_trans(easyPickImgAcqPose,p[0.0000,0.0000,-0.0000,0.0000,0.0000,0.0000]),a=1.3963,v=1.0472,t=0.000000,r=0.000000)
          easyPickAtImgAcq = True
        end
        easyPickPose = easyPickFuncTrigger(easyPickVisorId, easyPickSetJob, easyPickJobName, easyPickArmMounted)
      end
      # end: URCap Program Node
      # begin: URCap Program Node
      #   Source: SensoPart VISOR Robotic, 2.0.6, SensoPart Industriesensorik GmbH
      #   Type: Object Detected
      $ 2892 "Object Detected" "noBreak"
      if (visor_partsFound(easyPickVisorId) > 0):
        $ 2893 "Open Gripper" "noBreak"
        # begin: URCap Program Node
        #   Source: Robotiq_Grippers, 3.17.0.105337, Robotiq Inc.
        #   Type: Gripper
        $ 2894 "Gripper Open (1)" "noBreak"
        if not(gripper_connected[0]):
          popup("Gripper 1 must be connected to run this program.", "No connection", False, True, True)
        end
        if not(rq_is_gripper_activated("1")):
          popup("Gripper 1 is not activated. Go to Installation tab > Gripper to activate it and run the program again.", "Not activated", False, True, True)
        end
        rq_set_pos_spd_for(0, 77, 77, "1")
        rq_wait_pos_spe_for_request(0, 77, 77, "1")
        rq_go_to("1")
        rq_wait("1")
        # end: URCap Program Node
        $ 2895 "Set" "noBreak"
        set_tcp(p[0.0,0.0,0.161,3.1415,0.0,0.0])
        $ 2896 "Wait: 0.2" "noBreak"
        sleep(0.2)
        $ 2897 "Place on second weigh scale" "noBreak"
        $ 2898 "MoveJ" "noBreak"
        $ 2899 "Waypoint_1" "noBreak"
        movej(get_inverse_kin(Waypoint_1_p, qnear=Waypoint_1_q), a=1.3962634015954636, v=1.0471975511965976, r=0.1)
        $ 2900 "Waypoint_5" "noBreak"
        movej(get_inverse_kin(Waypoint_5_p, qnear=Waypoint_5_q), a=1.3962634015954636, v=1.0471975511965976)
        $ 2901 "read_db_data()" "noBreak"
        read_db_data()
        $ 2903 "Pick from B" "noBreak"
        $ 2904 "MoveL" "noBreak"
        $ 2906 "cont_B_safe" "noBreak"
        movel(cont_B_safe_p, a=1.2, v=0.25)
        $ 2907 "cont_B_prepick≔pose_trans(Cont_B_TCP, p[0,0,cent_edge/2,0,0,0])" "noBreak"
        global cont_B_prepick= pose_trans (Cont_B_TCP, p[0,0,cent_edge/2,0,0,0])
        $ 2908 "cont_B_otw" "noBreak"
        movel(cont_B_otw_p, a=1.2, v=0.25)
        $ 2910 "cont_B_pick≔pose_trans(cont_B_prepick, p[0,pick_2_base-d_cc,0,0,0,0])" "noBreak"
        global cont_B_pick= pose_trans (cont_B_prepick, p[0,pick_2_base-d_cc,0,0,0,0])
        $ 2911 "cont_B_pick" "noBreak"
        movel(cont_B_pick, a=0.2, v=0.1)
        # begin: URCap Program Node
        #   Source: Robotiq_Grippers, 3.17.0.105337, Robotiq Inc.
        #   Type: Gripper
        $ 2912 "Gripper Close (1)" "noBreak"
        if not(gripper_connected[0]):
          popup("Gripper 1 must be connected to run this program.", "No connection", False, True, True)
        end
        if not(rq_is_gripper_activated("1")):
          popup("Gripper 1 is not activated. Go to Installation tab > Gripper to activate it and run the program again.", "Not activated", False, True, True)
        end
        rq_set_pos_spd_for(255, 77, 51, "1")
        rq_wait_pos_spe_for_request(255, 77, 51, "1")
        rq_go_to("1")
        rq_wait("1")
        # end: URCap Program Node
        $ 2913 "cont_B_prepick" "noBreak"
        movel(cont_B_prepick, a=1.2, v=0.25, r=0.01)
        $ 2914 "Postions_otw" "noBreak"
        movel(Postions_otw_p, a=1.2, v=0.25)
        $ 2938 "Set" "noBreak"
        set_tcp(p[0.0,0.0,0.15052000000000001,3.1415,0.0,0.0])
        # begin: URCap Program Node
        #   Source: SensoPart VISOR Robotic, 2.0.6, SensoPart Industriesensorik GmbH
        #   Type: Approach Pose
        $ 2939 "Approach Pose" "noBreak"
        movej(pose_trans(easyPickPose,p[0.0000,0.0000,-0.0000,0.0000,0.0000,0.0000]),a=0.5236,v=0.4363,t=0.000000,r=0.000000)
        # end: URCap Program Node
        # begin: URCap Program Node
        #   Source: SensoPart VISOR Robotic, 2.0.6, SensoPart Industriesensorik GmbH
        #   Type: Target Pose
        $ 2940 "Target Pose" "noBreak"
        movel(pose_trans(easyPickPose,p[0.0000,0.0000,-0.0000,0.0000,0.0000,0.0000]),a=0.1000,v=0.0500,t=0.000000,r=0.000000)
        # end: URCap Program Node
        $ 2941 "Close Gripper" "noBreak"
        $ 2942 "container_place≔get_actual_tcp_pose()" "noBreak"
        global container_place= get_actual_tcp_pose ()
        $ 2943 "PoTS_place_abov≔pose_trans(container_place, p[0,0,cent_edge/2,0,0,0])" "noBreak"
        global PoTS_place_abov=pose_trans(container_place, p[0,0,cent_edge/2,0,0,0])
        $ 2945 "MoveL" "noBreak"
        $ 2946 "PoTS_place_abov" "noBreak"
        movel(PoTS_place_abov, a=0.5, v=0.05)
        $ 2947 "target_pose≔pose_trans(PoTS_place_abov, p[0,pick_2_base-d_cc,0,0,0,0])" "noBreak"
        global target_pose=pose_trans(PoTS_place_abov, p[0,pick_2_base-d_cc,0,0,0,0])
        $ 2948 "MoveL" "noBreak"
        $ 2949 "target_pose" "noBreak"
        movel(target_pose, a=0.3, v=0.05)
        # begin: URCap Program Node
        #   Source: Robotiq_Grippers, 3.17.0.105337, Robotiq Inc.
        #   Type: Gripper
        $ 2950 "Gripper Open (1)" "noBreak"
        if not(gripper_connected[0]):
          popup("Gripper 1 must be connected to run this program.", "No connection", False, True, True)
        end
        if not(rq_is_gripper_activated("1")):
          popup("Gripper 1 is not activated. Go to Installation tab > Gripper to activate it and run the program again.", "Not activated", False, True, True)
        end
        rq_set_pos_spd_for(0, 77, 77, "1")
        rq_wait_pos_spe_for_request(0, 77, 77, "1")
        rq_go_to("1")
        rq_wait("1")
        # end: URCap Program Node
        # begin: URCap Program Node
        #   Source: SensoPart VISOR Robotic, 2.0.6, SensoPart Industriesensorik GmbH
        #   Type: Exit Pose
        $ 2951 "Exit Pose" "noBreak"
        movel(pose_trans(easyPickPose,p[0.0000,0.0000,0.1000,0.0000,0.0000,0.0000]),a=0.5000,v=0.2500,t=0.000000,r=0.000000)
        # end: URCap Program Node
        easyPickObjTaken = True
      end
      # end: URCap Program Node
      # begin: URCap Program Node
      #   Source: SensoPart VISOR Robotic, 2.0.6, SensoPart Industriesensorik GmbH
      #   Type: No Object Detected
      $ 2952 "No Object Detected" "noBreak"
      if (visor_partsFound(easyPickVisorId) < 1):
        $ 2953 "Popup: No POTS detected" "noBreak"
        popup("No POTS detected", "Message", False, False, blocking=True)
        else:
      end
      # end: URCap Program Node
    end
    easyPickCount_7 = easyPickCount_7 + 1
    visor_easyPickUpdate(easyPickVisorId, "counter", easyPickCount_7)
    visor_easyPickSetIdent("133617", easyPickVisorId)
    # end: URCap Program Node
  end
  visorFuncEasyPick_316065()
  # end: URCap Program Node
  $ 2982 "MoveJ"
  $ 2983 "place_2_home" "breakAfter"
  movej(get_inverse_kin(place_2_home_p, qnear=place_2_home_q), a=1.3962634015954636, v=1.0471975511965976)
  elif (42 == switch_1):
    $ 2984 "Case 42"
  elif (43 == switch_1):
    $ 3746 "Case 43"
  elif (44 == switch_1):
    $ 3999 "Case 44"
    $ 4000 "Decap Container for recipe"
    $ 4002 "If powder_position ≟ 'Position1'"
    if (powder_position  ==  "Position1"):
      $ 4003 "MoveJ"
      $ 4004 "Postions_otw" "breakAfter"
      movej(get_inverse_kin(Postions_otw_p, qnear=Postions_otw_q), a=1.3962634015954636, v=1.0471975511965976, r=0.01)
      # begin: URCap Program Node
      #   Source: Robotiq_Grippers, 3.17.0.105337, Robotiq Inc.
      #   Type: Gripper
      $ 4005 "Gripper Open (1)"
      if not(gripper_connected[0]):
        popup("Gripper 1 must be connected to run this program.", "No connection", False, True, True)
      end
      if not(rq_is_gripper_activated("1")):
        popup("Gripper 1 is not activated. Go to Installation tab > Gripper to activate it and run the program again.", "Not activated", False, True, True)
      end
      rq_set_pos_spd_for(0, 127, 77, "1")
      rq_wait_pos_spe_for_request(0, 127, 77, "1")
      rq_go_to("1")
      rq_wait("1")
      # end: URCap Program Node
      $ 4006 "MoveL"
      $ 4007 "PosA_up" "breakAfter"
      movel(PosA_up_p, a=1.2, v=0.25)
      $ 4008 "PosA_pick" "breakAfter"
      movel(PosA_pick_p, a=1.2, v=0.25)
      # begin: URCap Program Node
      #   Source: Robotiq_Grippers, 3.17.0.105337, Robotiq Inc.
      #   Type: Gripper
      $ 4009 "Gripper Close (1)"
      if not(gripper_connected[0]):
        popup("Gripper 1 must be connected to run this program.", "No connection", False, True, True)
      end
      if not(rq_is_gripper_activated("1")):
        popup("Gripper 1 is not activated. Go to Installation tab > Gripper to activate it and run the program again.", "Not activated", False, True, True)
      end
      rq_set_pos_spd_for(255, 127, 77, "1")
      rq_wait_pos_spe_for_request(255, 127, 77, "1")
      rq_go_to("1")
      rq_wait("1")
      # end: URCap Program Node
      $ 4010 "PosA_up" "breakAfter"
      movel(PosA_up_p, a=0.3, v=0.04)
      $ 4011 "Postions_otw" "breakAfter"
      movel(Postions_otw_p, a=1.2, v=0.25, r=0.01)
    else:
      $ 4012 "ElseIf powder_position≟'Position2'"
      if (powder_position == "Position2"):
        $ 4013 "MoveJ"
        $ 4014 "Postions_otw" "breakAfter"
        movej(get_inverse_kin(Postions_otw_p, qnear=Postions_otw_q), a=1.3962634015954636, v=1.0471975511965976, r=0.01)
        # begin: URCap Program Node
        #   Source: Robotiq_Grippers, 3.17.0.105337, Robotiq Inc.
        #   Type: Gripper
        $ 4015 "Gripper Open (1)"
        if not(gripper_connected[0]):
          popup("Gripper 1 must be connected to run this program.", "No connection", False, True, True)
        end
        if not(rq_is_gripper_activated("1")):
          popup("Gripper 1 is not activated. Go to Installation tab > Gripper to activate it and run the program again.", "Not activated", False, True, True)
        end
        rq_set_pos_spd_for(0, 127, 77, "1")
        rq_wait_pos_spe_for_request(0, 127, 77, "1")
        rq_go_to("1")
        rq_wait("1")
        # end: URCap Program Node
        $ 4016 "MoveL"
        $ 4017 "PosB_up" "breakAfter"
        movel(PosB_up_p, a=1.2, v=0.25, r=0.01)
        $ 4018 "PosB_pick" "breakAfter"
        movel(PosB_pick_p, a=1.2, v=0.25)
        # begin: URCap Program Node
        #   Source: Robotiq_Grippers, 3.17.0.105337, Robotiq Inc.
        #   Type: Gripper
        $ 4019 "Gripper Close (1)"
        if not(gripper_connected[0]):
          popup("Gripper 1 must be connected to run this program.", "No connection", False, True, True)
        end
        if not(rq_is_gripper_activated("1")):
          popup("Gripper 1 is not activated. Go to Installation tab > Gripper to activate it and run the program again.", "Not activated", False, True, True)
        end
        rq_set_pos_spd_for(255, 127, 77, "1")
        rq_wait_pos_spe_for_request(255, 127, 77, "1")
        rq_go_to("1")
        rq_wait("1")
        # end: URCap Program Node
        $ 4020 "PosB_up" "breakAfter"
        movel(PosB_up_p, a=0.4, v=0.05)
        $ 4021 "Postions_otw" "breakAfter"
        movel(Postions_otw_p, a=1.2, v=0.25)
      else:
        $ 4022 "ElseIf powder_position≟'Position3'"
        if (powder_position == "Position3"):
          $ 4023 "MoveJ"
          $ 4024 "Postions_otw" "breakAfter"
          movej(get_inverse_kin(Postions_otw_p, qnear=Postions_otw_q), a=1.3962634015954636, v=1.0471975511965976, r=0.01)
          # begin: URCap Program Node
          #   Source: Robotiq_Grippers, 3.17.0.105337, Robotiq Inc.
          #   Type: Gripper
          $ 4025 "Gripper Open (1)"
          if not(gripper_connected[0]):
            popup("Gripper 1 must be connected to run this program.", "No connection", False, True, True)
          end
          if not(rq_is_gripper_activated("1")):
            popup("Gripper 1 is not activated. Go to Installation tab > Gripper to activate it and run the program again.", "Not activated", False, True, True)
          end
          rq_set_pos_spd_for(0, 127, 77, "1")
          rq_wait_pos_spe_for_request(0, 127, 77, "1")
          rq_go_to("1")
          rq_wait("1")
          # end: URCap Program Node
          $ 4026 "MoveL"
          $ 4027 "PosC_up" "breakAfter"
          movel(PosC_up_p, a=1.2, v=0.25, r=0.01)
          $ 4028 "PosC_pick" "breakAfter"
          movel(PosC_pick_p, a=1.2, v=0.25)
          # begin: URCap Program Node
          #   Source: Robotiq_Grippers, 3.17.0.105337, Robotiq Inc.
          #   Type: Gripper
          $ 4029 "Gripper Close (1)"
          if not(gripper_connected[0]):
            popup("Gripper 1 must be connected to run this program.", "No connection", False, True, True)
          end
          if not(rq_is_gripper_activated("1")):
            popup("Gripper 1 is not activated. Go to Installation tab > Gripper to activate it and run the program again.", "Not activated", False, True, True)
          end
          rq_set_pos_spd_for(255, 127, 77, "1")
          rq_wait_pos_spe_for_request(255, 127, 77, "1")
          rq_go_to("1")
          rq_wait("1")
          # end: URCap Program Node
          $ 4030 "PosC_up" "breakAfter"
          movel(PosC_up_p, a=0.5, v=0.05)
        end
      end
    end
    $ 4031 "MoveJ"
    $ 4032 "Pow_decap_up" "breakAfter"
    movej(get_inverse_kin(Pow_decap_up_p, qnear=Pow_decap_up_q), a=1.3962634015954636, v=1.0471975511965976)
    $ 4033 "Set GRP_3F_Open=On"
    set_standard_digital_out(5, True)
    $ 4034 "Wait: 0.5"
    sleep(0.5)
    $ 4035 "MoveL"
    $ 4036 "pow_decap_place" "breakAfter"
    movel(pow_decap_place_p, a=0.5, v=0.05)
    $ 4037 "Set GRP_3F_Open=Off"
    set_standard_digital_out(5, False)
    $ 4038 "Wait: 0.5"
    sleep(0.5)
    # begin: URCap Program Node
    #   Source: Robotiq_Grippers, 3.17.0.105337, Robotiq Inc.
    #   Type: Gripper
    $ 4039 "Gripper Open (1)"
    if not(gripper_connected[0]):
      popup("Gripper 1 must be connected to run this program.", "No connection", False, True, True)
    end
    if not(rq_is_gripper_activated("1")):
      popup("Gripper 1 is not activated. Go to Installation tab > Gripper to activate it and run the program again.", "Not activated", False, True, True)
    end
    rq_set_pos_spd_for(0, 255, 77, "1")
    rq_wait_pos_spe_for_request(0, 255, 77, "1")
    rq_go_to("1")
    rq_wait("1")
    # end: URCap Program Node
    $ 4040 "MoveL"
    $ 4041 "Pow_decap_up" "breakAfter"
    movel(Pow_decap_up_p, a=1.2, v=0.25)
    $ 4042 "Postions_otw" "breakAfter"
    movel(Postions_otw_p, a=1.2, v=0.25)
    $ 4043 "Home (Safe)"
    movej([-1.2302089344500047, -1.2969853503591224, -1.875639182904262, -1.539621866126728, 1.5731943360401213, -2.80099559440227], a=1.3962634015954636, v=1.0471975511965976)
    $ 4044 "MoveL"
    $ 4045 "Decap_above" "breakAfter"
    movel(Decap_above_p, a=1.2, v=0.25)
    $ 4046 "Decapp" "breakAfter"
    movel(Decapp_p, a=1.2, v=0.25)
    # begin: URCap Program Node
    #   Source: Robotiq_Grippers, 3.17.0.105337, Robotiq Inc.
    #   Type: Gripper
    $ 4047 "Gripper Close (1)"
    if not(gripper_connected[0]):
      popup("Gripper 1 must be connected to run this program.", "No connection", False, True, True)
    end
    if not(rq_is_gripper_activated("1")):
      popup("Gripper 1 is not activated. Go to Installation tab > Gripper to activate it and run the program again.", "Not activated", False, True, True)
    end
    rq_set_pos_spd_for(255, 128, 77, "1")
    rq_wait_pos_spe_for_request(255, 128, 77, "1")
    rq_go_to("1")
    rq_wait("1")
    # end: URCap Program Node
    $ 4048 "Decap"
    $ 4049 "Action_Info≔'decapping'"
    global Action_Info="decapping"
    $ 4050 "Set GRP_3F_Enable=On"
    set_standard_digital_out(4, True)
    $ 4051 "Set GRP_3F_Decap=On"
    set_standard_digital_out(3, True)
    $ 4052 "Force"
    sleep(0.02)
    zero_ftsensor()
    force_mode(p[0.0,0.0,0.0,0.0,0.0,0.0], [0, 0, 1, 0, 0, 0], [0.0, 0.0, 2.0, 0.0, 0.0, 0.0], 2, [0.1, 0.1, 5.0E-4, 0.3490658503988659, 0.3490658503988659, 0.3490658503988659])
    $ 4053 "check_decapping(offset=0.010, timeout=4.5, abort=CMD_Hold)" "noBreak"
    check_decapping(offset=0.010, timeout=4.5, abort=CMD_Hold)
    end_force_mode()
    stopl(5.0)
    $ 4054 "Set GRP_3F_Decap=Off"
    set_standard_digital_out(3, False)
    $ 4055 "Set GRP_3F_Enable=Off"
    set_standard_digital_out(4, False)
    $ 4056 "MoveL"
    $ 4057 "Decap_above" "breakAfter"
    movel(Decap_above_p, a=1.2, v=0.25)
    $ 4058 "Cap_above" "breakAfter"
    movel(Cap_above_p, a=1.2, v=0.25, r=0.05)
    $ 4059 "Cap_place" "breakAfter"
    movel(Cap_place_p, a=1.2, v=0.25)
    # begin: URCap Program Node
    #   Source: Robotiq_Grippers, 3.17.0.105337, Robotiq Inc.
    #   Type: Gripper
    $ 4060 "Gripper Move39mm (1)"
    if not(gripper_connected[0]):
      popup("Gripper 1 must be connected to run this program.", "No connection", False, True, True)
    end
    if not(rq_is_gripper_activated("1")):
      popup("Gripper 1 is not activated. Go to Installation tab > Gripper to activate it and run the program again.", "Not activated", False, True, True)
    end
    rq_set_pos_spd_for(67, 77, 77, "1")
    rq_wait_pos_spe_for_request(67, 77, 77, "1")
    rq_go_to("1")
    rq_wait("1")
    # end: URCap Program Node
    $ 4061 "Cap_above" "breakAfter"
    movel(Cap_above_p, a=1.2, v=0.25, r=0.05)
    $ 4062 "Home (Safe)"
    movej([-1.2302089344500047, -1.2969853503591224, -1.875639182904262, -1.539621866126728, 1.5731943360401213, -2.80099559440227], a=1.3962634015954636, v=1.0471975511965976)
  elif (45 == switch_1):
    $ 4063 "Case 45"
    $ 4064 "Place the decapped container- recipe"
    $ 4065 "tilt_to_home()"
    tilt_to_home()
    # begin: URCap Program Node
    #   Source: SensoPart VISOR Robotic, 2.0.6, SensoPart Industriesensorik GmbH
    #   Type: VISOR Robotic App
    $ 4067 "VISOR Easy Pick"
    def visorFuncEasyPick_0d9b38():
      # begin: URCap Program Node
      #   Source: SensoPart VISOR Robotic, 2.0.6, SensoPart Industriesensorik GmbH
      #   Type: Easy Pick Setup
      $ 4068 "# 1 Setup" "noBreak"
      local easyPickVisorId = 1
      local easyPickArmMounted = True
      local easyPickSetJob = True
      local easyPickJobName = "PoTS"
      local easyPickAtImgAcq = False
      local easyPickImgAcqPose = Trigger
      # end: URCap Program Node
      # begin: URCap Program Node
      #   Source: SensoPart VISOR Robotic, 2.0.6, SensoPart Industriesensorik GmbH
      #   Type: Process
      $ 4069 "Process" "noBreak"
      local easyPickObjTaken = False
      local easyPickTrigger = False
      local easyPickPoseIdx = 0
      local easyPickPose = p[0,0,0,0,0,0]
      def easyPickFuncTrigger(visorId, setJob, jobName, arm):
      if (setJob):
        visor_changeJob(visorId, jobName, 6000)
      end
      if (arm):
        visor_trigger(visorId, 6000, "arm")
      else:
        visor_trigger(visorId, 6000)
      end
      global easyPickParts_7=visor_partsFound(visorId)
      visor_easyPickUpdate(visorId, "parts", visor_partsFound(visorId))
      return visor_getPose3d(visorId, 0)
    end
    while (not easyPickObjTaken):
      easyPickTrigger = (easyPickCount_7 >= visor_partsFound(easyPickVisorId)) or (easyPickCount_7 > 9) or (not visor_easyPickCheckIdent("a9cf93", easyPickVisorId))
      if (easyPickTrigger):
        easyPickCount_7 = 0
      end
      easyPickPoseIdx = easyPickCount_7
      easyPickPose = visor_getPose3d(easyPickVisorId, easyPickPoseIdx)
      visor_easyPickUpdate(easyPickVisorId, "counter", easyPickPoseIdx)
      # begin: URCap Program Node
      #   Source: SensoPart VISOR Robotic, 2.0.6, SensoPart Industriesensorik GmbH
      #   Type: Image Acquisition Pose
      $ 4070 "Image Acquisition Pose" "noBreak"
      if (easyPickTrigger):
        if (not easyPickAtImgAcq):
          movej(pose_trans(easyPickImgAcqPose,p[0.0000,0.0000,-0.0000,0.0000,0.0000,0.0000]),a=1.3963,v=1.0472,t=0.000000,r=0.000000)
          easyPickAtImgAcq = True
        end
        easyPickPose = easyPickFuncTrigger(easyPickVisorId, easyPickSetJob, easyPickJobName, easyPickArmMounted)
      end
      # end: URCap Program Node
      # begin: URCap Program Node
      #   Source: SensoPart VISOR Robotic, 2.0.6, SensoPart Industriesensorik GmbH
      #   Type: Object Detected
      $ 4071 "Object Detected" "noBreak"
      if (visor_partsFound(easyPickVisorId) > 0):
        $ 4072 "Open Gripper" "noBreak"
        # begin: URCap Program Node
        #   Source: Robotiq_Grippers, 3.17.0.105337, Robotiq Inc.
        #   Type: Gripper
        $ 4073 "Gripper Open (1)" "noBreak"
        if not(gripper_connected[0]):
          popup("Gripper 1 must be connected to run this program.", "No connection", False, True, True)
        end
        if not(rq_is_gripper_activated("1")):
          popup("Gripper 1 is not activated. Go to Installation tab > Gripper to activate it and run the program again.", "Not activated", False, True, True)
        end
        rq_set_pos_spd_for(0, 77, 77, "1")
        rq_wait_pos_spe_for_request(0, 77, 77, "1")
        rq_go_to("1")
        rq_wait("1")
        # end: URCap Program Node
        $ 4074 "MoveL" "noBreak"
        $ 4075 "OP_PowderA2" "noBreak"
        movel(OP_PowderA2_p, a=1.2, v=0.25)
        $ 4076 "Decap_up" "noBreak"
        movel(Decap_up_p, a=1.2, v=0.25)
        $ 4077 "Decap_pick" "noBreak"
        movel(Decap_pick_p, a=1.2, v=0.25)
        # begin: URCap Program Node
        #   Source: Robotiq_Grippers, 3.17.0.105337, Robotiq Inc.
        #   Type: Gripper
        $ 4078 "Gripper Close (1)" "noBreak"
        if not(gripper_connected[0]):
          popup("Gripper 1 must be connected to run this program.", "No connection", False, True, True)
        end
        if not(rq_is_gripper_activated("1")):
          popup("Gripper 1 is not activated. Go to Installation tab > Gripper to activate it and run the program again.", "Not activated", False, True, True)
        end
        rq_set_pos_spd_for(255, 77, 77, "1")
        rq_wait_pos_spe_for_request(255, 77, 77, "1")
        rq_go_to("1")
        rq_wait("1")
        # end: URCap Program Node
        $ 4079 "Wait: 0.5" "noBreak"
        sleep(0.5)
        $ 4080 "Set GRP_3F_Open=On" "noBreak"
        set_standard_digital_out(5, True)
        $ 4081 "Decap_up" "noBreak"
        movel(Decap_up_p, a=0.5, v=0.1)
        $ 4083 "Op_PowA_wP" "noBreak"
        movel(Op_PowA_wP_p, a=1.2, v=0.25)
        # begin: URCap Program Node
        #   Source: SensoPart VISOR Robotic, 2.0.6, SensoPart Industriesensorik GmbH
        #   Type: Approach Pose
        $ 4084 "Approach Pose" "noBreak"
        movej(pose_trans(easyPickPose,p[0.0000,0.0000,-0.0000,0.0000,0.0000,0.0000]),a=0.5236,v=0.4363,t=0.000000,r=0.000000)
        # end: URCap Program Node
        # begin: URCap Program Node
        #   Source: SensoPart VISOR Robotic, 2.0.6, SensoPart Industriesensorik GmbH
        #   Type: Target Pose
        $ 4085 "Target Pose" "noBreak"
        movel(pose_trans(easyPickPose,p[0.0000,0.0000,-0.0000,0.0000,0.0000,0.0000]),a=0.1000,v=0.0500,t=0.000000,r=0.000000)
        # end: URCap Program Node
        $ 4086 "Close Gripper" "noBreak"
        $ 4087 "container_place≔get_actual_tcp_pose()" "noBreak"
        global container_place= get_actual_tcp_pose ()
        $ 4088 "target_pose≔pose_add(container_place, p[0,0,-0.12,0,0,0])" "noBreak"
        global target_pose=pose_add(container_place, p[0,0,-0.12,0,0,0])
        $ 4089 "MoveL" "noBreak"
        $ 4090 "target_pose" "noBreak"
        movel(target_pose, a=0.3, v=0.05)
        # begin: URCap Program Node
        #   Source: Robotiq_Grippers, 3.17.0.105337, Robotiq Inc.
        #   Type: Gripper
        $ 4091 "Gripper Open (1)" "noBreak"
        if not(gripper_connected[0]):
          popup("Gripper 1 must be connected to run this program.", "No connection", False, True, True)
        end
        if not(rq_is_gripper_activated("1")):
          popup("Gripper 1 is not activated. Go to Installation tab > Gripper to activate it and run the program again.", "Not activated", False, True, True)
        end
        rq_set_pos_spd_for(0, 77, 77, "1")
        rq_wait_pos_spe_for_request(0, 77, 77, "1")
        rq_go_to("1")
        rq_wait("1")
        # end: URCap Program Node
        # begin: URCap Program Node
        #   Source: SensoPart VISOR Robotic, 2.0.6, SensoPart Industriesensorik GmbH
        #   Type: Exit Pose
        $ 4092 "Exit Pose" "noBreak"
        movel(pose_trans(easyPickPose,p[0.0000,0.0000,-0.0000,0.0000,0.0000,0.0000]),a=0.5000,v=0.2500,t=0.000000,r=0.000000)
        # end: URCap Program Node
        easyPickObjTaken = True
      end
      # end: URCap Program Node
      # begin: URCap Program Node
      #   Source: SensoPart VISOR Robotic, 2.0.6, SensoPart Industriesensorik GmbH
      #   Type: No Object Detected
      $ 4093 "No Object Detected" "noBreak"
      if (visor_partsFound(easyPickVisorId) < 1):
        $ 4094 "Popup: No weigh scale detected" "noBreak"
        popup("No weigh scale detected", "Message", False, False, blocking=True)
        else:
      end
      # end: URCap Program Node
    end
    easyPickCount_7 = easyPickCount_7 + 1
    visor_easyPickUpdate(easyPickVisorId, "counter", easyPickCount_7)
    visor_easyPickSetIdent("a9cf93", easyPickVisorId)
    # end: URCap Program Node
  end
  visorFuncEasyPick_0d9b38()
  # end: URCap Program Node
  $ 4095 "place_pose≔get_actual_tcp_pose()"
  global place_pose= get_actual_tcp_pose ()
  $ 4096 "center_pose()"
  center_pose()
  $ 4098 "MoveJ"
  $ 4099 "Waypoint_1" "breakAfter"
  movej(get_inverse_kin(Waypoint_1_p, qnear=Waypoint_1_q), a=1.3962634015954636, v=1.0471975511965976)
  elif (46 == switch_1):
    $ 4100 "Case 46"
  elif (47 == switch_1):
    $ 4390 "Case 47"
  elif (48 == switch_1):
    $ 4445 "Case 48"
  elif (49 == switch_1):
    $ 4463 "Case 49"
  elif (50 == switch_1):
    $ 4481 "Case 50"
    $ 4482 "Emptying powder container"
    $ 4483 "Dosing untill empty"
    $ 4484 "send_target_info()"
    send_target_info()
    $ 4485 "zero_scale()"
    zero_scale()
    $ 4486 "prev_spat≔''"
    global prev_spat=""
    $ 4487 "spatula≔''"
    global spatula=""
    $ 4488 "send_powder_info()"
    send_powder_info()
    $ 4489 "Set AO[0]=0.0"
    set_standard_analog_out(0, 0.0)
    $ 4490 "Wait: 0.2"
    sleep(0.2)
    $ 4491 "reach pots decapping pose"
    # begin: URCap Program Node
    #   Source: SensoPart VISOR Robotic, 2.0.6, SensoPart Industriesensorik GmbH
    #   Type: VISOR Robotic App
    $ 4497 "VISOR Easy Pick"
    def visorFuncEasyPick_971e99():
      # begin: URCap Program Node
      #   Source: SensoPart VISOR Robotic, 2.0.6, SensoPart Industriesensorik GmbH
      #   Type: Easy Pick Setup
      $ 4498 "# 1 Setup" "noBreak"
      local easyPickVisorId = 1
      local easyPickArmMounted = True
      local easyPickSetJob = True
      local easyPickJobName = "Weight_scale"
      local easyPickAtImgAcq = False
      local easyPickImgAcqPose = Trigger
      # end: URCap Program Node
      # begin: URCap Program Node
      #   Source: SensoPart VISOR Robotic, 2.0.6, SensoPart Industriesensorik GmbH
      #   Type: Process
      $ 4499 "Process" "noBreak"
      local easyPickObjTaken = False
      local easyPickTrigger = False
      local easyPickPoseIdx = 0
      local easyPickPose = p[0,0,0,0,0,0]
      def easyPickFuncTrigger(visorId, setJob, jobName, arm):
      if (setJob):
        visor_changeJob(visorId, jobName, 6000)
      end
      if (arm):
        visor_trigger(visorId, 6000, "arm")
      else:
        visor_trigger(visorId, 6000)
      end
      global easyPickParts_4=visor_partsFound(visorId)
      visor_easyPickUpdate(visorId, "parts", visor_partsFound(visorId))
      return visor_getPose3d(visorId, 0)
    end
    while (not easyPickObjTaken):
      easyPickTrigger = (easyPickCount_4 >= visor_partsFound(easyPickVisorId)) or (easyPickCount_4 > 9) or (not visor_easyPickCheckIdent("20fd05", easyPickVisorId))
      if (easyPickTrigger):
        easyPickCount_4 = 0
      end
      easyPickPoseIdx = easyPickCount_4
      easyPickPose = visor_getPose3d(easyPickVisorId, easyPickPoseIdx)
      visor_easyPickUpdate(easyPickVisorId, "counter", easyPickPoseIdx)
      # begin: URCap Program Node
      #   Source: SensoPart VISOR Robotic, 2.0.6, SensoPart Industriesensorik GmbH
      #   Type: Image Acquisition Pose
      $ 4500 "Image Acquisition Pose" "noBreak"
      if (easyPickTrigger):
        if (not easyPickAtImgAcq):
          movej(pose_trans(easyPickImgAcqPose,p[0.0000,0.0000,-0.0000,0.0000,0.0000,0.0000]),a=1.3963,v=1.0472,t=0.000000,r=0.000000)
          easyPickAtImgAcq = True
        end
        easyPickPose = easyPickFuncTrigger(easyPickVisorId, easyPickSetJob, easyPickJobName, easyPickArmMounted)
      end
      # end: URCap Program Node
      # begin: URCap Program Node
      #   Source: SensoPart VISOR Robotic, 2.0.6, SensoPart Industriesensorik GmbH
      #   Type: Object Detected
      $ 4501 "Object Detected" "noBreak"
      if (visor_partsFound(easyPickVisorId) > 0):
        $ 4502 "Open Gripper" "noBreak"
        $ 4503 "weight_value≔get_weight()" "noBreak"
        global weight_value=get_weight()
        $ 4504 "Wait: 1.0" "noBreak"
        sleep(1.0)
        $ 4505 "diff≔target_weight-weight_value" "noBreak"
        global diff=target_weight-weight_value
        $ 4506 "compute_level_percent(W_now, weight_value)" "noBreak"
        compute_level_percent(W_now, weight_value)
        $ 4507 "send_level_info()" "noBreak"
        send_level_info()
        $ 4508 "spatula≔select_spatula(Flowability, level, diff, bulk_density, mouth_d)" "noBreak"
        global spatula=select_spatula(Flowability, level, diff, bulk_density, mouth_d)
        $ 4509 "Wait: 0.2" "noBreak"
        sleep(0.2)
        $ 4510 "send_spatula_info()" "noBreak"
        send_spatula_info()
        $ 4511 "If spatula ≟ 'spatula_L'" "noBreak"
        if (spatula  ==  "spatula_L"):
          $ 4512 "MoveJ" "noBreak"
          $ 4513 "Spatula_otw" "noBreak"
          movej(get_inverse_kin(Spatula_otw_p, qnear=Spatula_otw_q), a=1.3962634015954636, v=1.0471975511965976)
          $ 4514 "pick_spat_L_abv" "noBreak"
          movej(get_inverse_kin(pick_spat_L_abv_p, qnear=pick_spat_L_abv_q), a=1.3962634015954636, v=1.0471975511965976)
          $ 4515 "MoveL" "noBreak"
          $ 4516 "spat_L_pick" "noBreak"
          movel(spat_L_pick_p, a=1.2, v=0.25)
          # begin: URCap Program Node
          #   Source: Robotiq_Grippers, 3.17.0.105337, Robotiq Inc.
          #   Type: Gripper
          $ 4517 "Gripper Close (1)" "noBreak"
          if not(gripper_connected[0]):
            popup("Gripper 1 must be connected to run this program.", "No connection", False, True, True)
          end
          if not(rq_is_gripper_activated("1")):
            popup("Gripper 1 is not activated. Go to Installation tab > Gripper to activate it and run the program again.", "Not activated", False, True, True)
          end
          rq_set_pos_spd_for(255, 0, 77, "1")
          rq_wait_pos_spe_for_request(255, 0, 77, "1")
          rq_go_to("1")
          rq_wait("1")
          # end: URCap Program Node
          $ 4518 "spat_L_lift" "noBreak"
          movel(spat_L_lift_p, a=1.2, v=0.25, r=0.01)
          $ 4519 "spat_L_side" "noBreak"
          movel(spat_L_side_p, a=1.2, v=0.25, r=0.01)
          $ 4520 "spat_L_up" "noBreak"
          movel(spat_L_up_p, a=1.2, v=0.25, r=0.05)
          $ 4521 "MoveJ" "noBreak"
          $ 4522 "Spatula_otw" "noBreak"
          movej(get_inverse_kin(Spatula_otw_p, qnear=Spatula_otw_q), a=1.3962634015954636, v=1.0471975511965976)
        else:
          $ 4523 "ElseIf spatula ≟'spatula_M'" "noBreak"
          if (spatula  == "spatula_M"):
            $ 4524 "MoveJ" "noBreak"
            $ 4525 "Spatula_otw" "noBreak"
            movej(get_inverse_kin(Spatula_otw_p, qnear=Spatula_otw_q), a=1.3962634015954636, v=1.0471975511965976)
            $ 4526 "spat_M_up" "noBreak"
